	// xBusy не покрывает удерживаемый запрос и завершение Disable.
	// Занятость другого магазина/станка сама по себе не запрещает правку инвентаря.
	xTwinRobotOperation := GVL_MAGAZINE.astPartStatus[uiTwin].xBusy
		OR GVL_MAGAZINE.astPartStatus[uiTwin].xDisablePending
		OR GVL_MAGAZINE.astAutoCommand[uiTwin].xExecute
		OR GVL_MAGAZINE.astCommand[uiTwin].xExecute
		OR ((GVL_ROBOT.Status.xBusy OR xMotionBusy)
			AND (GVL_ROBOT.Status.uiMagazineContext = uiTwin))
		OR ((GVL_CELL_MANAGER.Status.uiActiveMagazine = uiTwin)
			AND ((GVL_CELL_MANAGER.Diag.eState = E_CELL_STATE.MAGAZINE)
				OR (GVL_CELL_MANAGER.Diag.eState = E_CELL_STATE.RELEASE_MAGAZINE)));
	// Для обмена важна занятость только этого магазина. Точка и состояние
	// интерфейса робота после инициализации могут быть неизвестны.
	xTwinRobotSwapWindow := NOT xTwinRobotOperation;
	xTwinOtherLoaded := FALSE;
	IF (GVL_TWO_PALLET.astStatus[uiTwin].uiRobotPallet >= UINT#1)
		AND (GVL_TWO_PALLET.astStatus[uiTwin].uiRobotPallet <= UINT#2) THEN
		uiTwinPallet := UINT#3 - GVL_TWO_PALLET.astStatus[uiTwin].uiRobotPallet;
		xTwinOtherLoaded := GVL_TWO_PALLET.astStore[uiTwin].axLoaded[uiTwinPallet];
	END_IF;
	// Finished удерживает цикл в ожидании даже до подтверждения загрузки второй палеты.
	// Подтверждение, разрешение автообмена и готовность зоны отдельно разрешают движение.
	axTwinAutoSwapPending[uiTwin] := (GVL_TWO_PALLET.uiMode = UINT#1)
		AND GVL_CELL_MANAGER.Status.xRunning
		AND NOT GVL_CELL_MANAGER.Status.xStopPending
		AND NOT GVL_CELL_CONTROL.xStop
		AND NOT GVL_CELL_CONTROL.xManual
		AND GVL_MAGAZINE.astPartStatus[uiTwin].xFinished
		AND NOT astTwinCommand[uiTwin].xDisable
		AND NOT astTwinCommand[uiTwin].xStop;
	uiTwinRobotPalletBefore := GVL_TWO_PALLET.astStatus[uiTwin].uiRobotPallet;
	TWIN[uiTwin](
		xSelected := GVL_TWO_PALLET.uiMode = 1,
		xManual := GVL_CELL_CONTROL.xManual AND NOT GVL_CELL_MANAGER.Status.xRunning,
		xSafe := CELL_SAFETY.Status.xReady AND NOT GVL_CELL_CONTROL.xGlobalError AND NOT GVL_HMI.xIoEmergencyStopActive
			AND CELL_SAFETY.astEnclosureDoorStatus[uiTwin * 2 - 1].xLocked
			AND CELL_SAFETY.astEnclosureDoorStatus[uiTwin * 2].xLocked
			AND NOT CELL_SAFETY.astEnclosureDoorStatus[uiTwin * 2 - 1].xUnlockOutput
			AND NOT CELL_SAFETY.astEnclosureDoorStatus[uiTwin * 2].xUnlockOutput,
		xRobotSwapWindow := xTwinRobotSwapWindow,
		xRobotOperation := xTwinRobotOperation,
		xPointsConfigured := axMagazinePointsReady[uiTwin],
		xRobotGeometryReady := NOT GVL_HMI.xModbusMode AND axMagazinePointsReady[uiTwin],
		xRobotMagazineReady := GVL_MAGAZINE.astPartStatus[uiTwin].xEnableCheckNoError
			AND GVL_MAGAZINE.astPartStatus[uiTwin].xEnableCheckGeometry,
		xConnection := xHmiConnectionAlive,
		xStopRequest := GVL_CELL_CONTROL.xStop OR xIoManualActive OR GVL_HMI.astMagazineCommand[uiTwin].xStop OR GVL_TWO_PALLET.xModeChanged,
		xAutoSwap := axTwinAutoSwapPending[uiTwin] AND xTwinAutoSwapEnabled AND xTwinOtherLoaded,
		xOtherLoaded := xTwinOtherLoaded,
		xActivePalletEditAllowed := NOT xTwinRobotOperation,
		xConfigurationChanged := axTwinConfigurationChanged[uiTwin],
        xIoPneumaticOverride := axIoMagazineInvalidated[uiTwin],
		xExternalCommandRejected := axTwinExternalCommandRejected[uiTwin],
		Command := astTwinCommand[uiTwin],
		Config := GVL_TWO_PALLET.astActiveConfig[uiTwin], Input := GVL_TWO_PALLET.astInput[uiTwin],
		Status => GVL_TWO_PALLET.astStatus[uiTwin],
		Diag => GVL_TWO_PALLET.astDiag[uiTwin],
		Error => GVL_TWO_PALLET.astError[uiTwin],
		Output => GVL_TWO_PALLET.astOutput[uiTwin]);
    axIoMagazineInvalidated[uiTwin] := FALSE;
	// Блокировка относится только к этому магазину и удерживается до полного
	// окончания механического обмена, включая последний скан Completed.
	axTwinMagazineExchangeInProgress[uiTwin] := GVL_TWO_PALLET.astStatus[uiTwin].xBusy
		OR GVL_TWO_PALLET.astStatus[uiTwin].xCompleted;
	GVL_TWO_PALLET.astStatus[uiTwin].xAutoSwapEnabled := xTwinAutoSwapEnabled;
	// После Stop/Disable или аварии ожидание обмена не удерживает планировщик.
	axTwinAutoSwapPending[uiTwin] := axTwinAutoSwapPending[uiTwin]
		AND NOT GVL_TWO_PALLET.astStatus[uiTwin].xError;
	axTwinConfigurationChanged[uiTwin] := FALSE;
	axTwinExternalCommandRejected[uiTwin] := FALSE;
	IF GVL_TWO_PALLET.astOutput[uiTwin].xTeachOperator THEN
		IF GVL_CELL_SETTINGS.eTestEnvironment = E_CELL_TEST_ENVIRONMENT.SIMULATION THEN
			GVL_TWO_PALLET.astSimulationConfig[uiTwin].lrExchange := GVL_TWO_PALLET.astInput[uiTwin].lrPosition;
		ELSE
			GVL_TWO_PALLET.astConfig[uiTwin].lrExchange := GVL_TWO_PALLET.astInput[uiTwin].lrPosition;
		END_IF;
		axTwinConfigurationChanged[uiTwin] := TRUE;
	END_IF;
	IF GVL_TWO_PALLET.astOutput[uiTwin].xTeachWork THEN
		IF GVL_TWO_PALLET.astStatus[uiTwin].uiSelected = UINT#1 THEN
			IF GVL_CELL_SETTINGS.eTestEnvironment = E_CELL_TEST_ENVIRONMENT.SIMULATION THEN
				GVL_TWO_PALLET.astSimulationConfig[uiTwin].lrWorkP1 := GVL_TWO_PALLET.astInput[uiTwin].lrPosition;
			ELSE
				GVL_TWO_PALLET.astConfig[uiTwin].lrWorkP1 := GVL_TWO_PALLET.astInput[uiTwin].lrPosition;
			END_IF;
		ELSIF GVL_TWO_PALLET.astStatus[uiTwin].uiSelected = UINT#2 THEN
			IF GVL_CELL_SETTINGS.eTestEnvironment = E_CELL_TEST_ENVIRONMENT.SIMULATION THEN
				GVL_TWO_PALLET.astSimulationConfig[uiTwin].lrWorkP2 := GVL_TWO_PALLET.astInput[uiTwin].lrPosition;
			ELSE
				GVL_TWO_PALLET.astConfig[uiTwin].lrWorkP2 := GVL_TWO_PALLET.astInput[uiTwin].lrPosition;
			END_IF;
		END_IF;
		axTwinConfigurationChanged[uiTwin] := TRUE;
	END_IF;
	// RunCellControl ниже должен видеть запрет уже в скане начала обмена.
	IF GVL_TWO_PALLET.uiMode = 1 THEN
		GVL_MAGAZINE.astStatus[uiTwin].xReady := GVL_MAGAZINE.astPartStatus[uiTwin].xReady
			AND GVL_TWO_PALLET.astStatus[uiTwin].xReady;
		GVL_MAGAZINE.astStatus[uiTwin].xBusy := GVL_MAGAZINE.astPartStatus[uiTwin].xBusy
			OR GVL_TWO_PALLET.astStatus[uiTwin].xBusy;
		GVL_MAGAZINE.astStatus[uiTwin].xEnabled := GVL_TWO_PALLET.astStatus[uiTwin].xEnabled;
	END_IF;
	IF GVL_TWO_PALLET.astStatus[uiTwin].xCompleted THEN
		GVL_TWO_PALLET.astStore[uiTwin].axLoaded[1] := FALSE;
		GVL_TWO_PALLET.astStore[uiTwin].axLoaded[2] := FALSE;
		axMagazineInventoryChanged[uiTwin] := TRUE;
	END_IF;
	// Ручное восстановление может сменить учётную роль без команды обмена.
	IF uiTwinRobotPalletBefore <> GVL_TWO_PALLET.astStatus[uiTwin].uiRobotPallet THEN
		GVL_TWO_PALLET.astStore[uiTwin].axLoaded[1] := FALSE;
		GVL_TWO_PALLET.astStore[uiTwin].axLoaded[2] := FALSE;
		axMagazineInventoryChanged[uiTwin] := TRUE;
	END_IF;
	// Ручная смена расходует прежнее подтверждение уже при принятии команды.
	IF astTwinCommand[uiTwin].xSwap AND GVL_TWO_PALLET.astStatus[uiTwin].xCommandAccepted THEN
		GVL_TWO_PALLET.astStore[uiTwin].axLoaded[1] := FALSE;
		GVL_TWO_PALLET.astStore[uiTwin].axLoaded[2] := FALSE;
	END_IF;
	IF (uiTwinRequestResult = 2) AND (stTwinRequest.uiMagazine = uiTwin)
		AND (((stTwinRequest.uiCommand >= 1) AND (stTwinRequest.uiCommand <= 19))
			OR ((stTwinRequest.uiCommand >= 25) AND (stTwinRequest.uiCommand <= 32)))
		AND GVL_TWO_PALLET.astStatus[uiTwin].xCommandAccepted THEN uiTwinRequestResult := 1; END_IF;
END_FOR;

IF xTwinInventoryCommand THEN
	uiTwin := stTwinRequest.uiMagazine;
	uiTwinPallet := stTwinRequest.uiValue;
	IF stTwinRequest.uiCommand = UINT#24 THEN
		IF GVL_TWO_PALLET.astStatus[uiTwin].xConfigAllowed
			AND stTwinRequest.Config.xSignalPatternsConfigured
			AND TWIN[uiTwin].IsSignalConfigurationValid(
				uiP1Signals := stTwinRequest.Config.uiP1Signals,
				uiP2Signals := stTwinRequest.Config.uiP2Signals) THEN
			IF GVL_CELL_SETTINGS.eTestEnvironment = E_CELL_TEST_ENVIRONMENT.SIMULATION THEN
				GVL_TWO_PALLET.astSimulationConfig[uiTwin] := stTwinRequest.Config;
			ELSE
				GVL_TWO_PALLET.astConfig[uiTwin] := stTwinRequest.Config;
			END_IF;
			axTwinConfigurationChanged[uiTwin] := TRUE;
			uiTwinRequestResult := UINT#1;
		END_IF;
	ELSIF ((uiTwinPallet = 1) AND GVL_TWO_PALLET.astStatus[uiTwin].xEdit1Allowed)
		OR ((uiTwinPallet = 2) AND GVL_TWO_PALLET.astStatus[uiTwin].xEdit2Allowed) THEN
		CASE stTwinRequest.uiCommand OF
			20:
				IF GVL_TWO_PALLET.astStatus[uiTwin].xLoadAllowed
					AND (uiTwinPallet <> GVL_TWO_PALLET.astStatus[uiTwin].uiRobotPallet) THEN
					GVL_TWO_PALLET.astStore[uiTwin].axLoaded[uiTwinPallet] := TRUE;
					uiTwinRequestResult := 1;
				END_IF;
			21, 22:
				FOR uiTwinSlot := 1 TO 96 DO
					GVL_TWO_PALLET.astStore[uiTwin].astPallet[uiTwinPallet].aSlots[uiTwinSlot].xInPosition := stTwinRequest.uiCommand = 22;
					GVL_TWO_PALLET.astStore[uiTwin].astPallet[uiTwinPallet].aSlots[uiTwinSlot].eDetailType := E_DETAIL_TYPE.NONE;
					GVL_TWO_PALLET.astStore[uiTwin].astPallet[uiTwinPallet].aSlots[uiTwinSlot].uiProductType := 0;
					IF stTwinRequest.uiCommand = 22 THEN
						GVL_TWO_PALLET.astStore[uiTwin].astPallet[uiTwinPallet].aSlots[uiTwinSlot].eDetailType := E_DETAIL_TYPE.BLANK;
						GVL_TWO_PALLET.astStore[uiTwin].astPallet[uiTwinPallet].aSlots[uiTwinSlot].uiProductType := GVL_MULTI_TYPE.Config.auiSlotType[uiTwinSlot];
					END_IF;
				END_FOR;
				GVL_TWO_PALLET.astStore[uiTwin].axLoaded[uiTwinPallet] := FALSE; uiTwinRequestResult := 1;
			23:
				IF (stTwinRequest.uiSlot >= 1) AND (stTwinRequest.uiSlot <= 96) AND (stTwinRequest.uiContent <= 2)
					AND ((stTwinRequest.uiContent = 0) OR ((stTwinRequest.uiProductType >= 1) AND (stTwinRequest.uiProductType <= GVL_MULTI_TYPE.Config.uiTypeCount))) THEN
					uiTwinSlot := stTwinRequest.uiSlot;
					GVL_TWO_PALLET.astStore[uiTwin].astPallet[uiTwinPallet].aSlots[uiTwinSlot].xInPosition := stTwinRequest.uiContent <> 0;
					CASE stTwinRequest.uiContent OF
						0: GVL_TWO_PALLET.astStore[uiTwin].astPallet[uiTwinPallet].aSlots[uiTwinSlot].eDetailType := E_DETAIL_TYPE.NONE;
						1: GVL_TWO_PALLET.astStore[uiTwin].astPallet[uiTwinPallet].aSlots[uiTwinSlot].eDetailType := E_DETAIL_TYPE.BLANK;
						2: GVL_TWO_PALLET.astStore[uiTwin].astPallet[uiTwinPallet].aSlots[uiTwinSlot].eDetailType := E_DETAIL_TYPE.DETAIL;
					END_CASE;
					GVL_TWO_PALLET.astStore[uiTwin].astPallet[uiTwinPallet].aSlots[uiTwinSlot].uiProductType := stTwinRequest.uiProductType;
					GVL_TWO_PALLET.astStore[uiTwin].axLoaded[uiTwinPallet] := FALSE; uiTwinRequestResult := 1;
				END_IF;
		END_CASE;
		// Загрузка/редактирование палеты у оператора не отменяет завершение рабочей.
		IF (uiTwinRequestResult = UINT#1)
			AND (stTwinRequest.uiCommand >= UINT#21)
			AND (stTwinRequest.uiCommand <= UINT#23)
			AND (uiTwinPallet = GVL_TWO_PALLET.astStatus[uiTwin].uiRobotPallet) THEN
			axMagazineInventoryChanged[uiTwin] := TRUE;
		END_IF;
	END_IF;
END_IF;
IF uiTwinRequestResult <> 0 THEN
	GVL_HMI.uiTwinResult := uiTwinRequestResult;
	GVL_HMI.udiTwinAckSeq := udiTwinSnapshot;
	IF uiTwinRequestResult <> 1 THEN
		uiTwin := LIMIT(UINT#1, stTwinRequest.uiMagazine, UINT#2);
		// Команды механизма 1..19 и 25..28 уже формируют предупреждение внутри FB в этом же скане.
		IF GVL_TWO_PALLET.auiCommand[uiTwin] <> stTwinRequest.uiCommand THEN
			axTwinExternalCommandRejected[uiTwin] := TRUE;
		END_IF;
	END_IF;
END_IF;

GVL_CELL_SETTINGS.MagazineRows := 12;
GVL_CELL_SETTINGS.MagazineColumns := 10;
IF GVL_TWO_PALLET.uiMode = 1 THEN GVL_CELL_SETTINGS.MagazineRows := 12; GVL_CELL_SETTINGS.MagazineColumns := 8; END_IF;
GVL_HMI.MagazineRows := GVL_CELL_SETTINGS.MagazineRows;
GVL_HMI.MagazineColumns := GVL_CELL_SETTINGS.MagazineColumns;
FOR uiTwin := 1 TO 2 DO
	IF GVL_TWO_PALLET.uiMode = 1 THEN
		uiTwinPallet := GVL_TWO_PALLET.astStatus[uiTwin].uiRobotPallet;
		IF (uiTwinPallet < UINT#1) OR (uiTwinPallet > UINT#2) THEN
			uiTwinPallet := UINT#1;
		END_IF;
		GVL_DETAIL.astMagazine[uiTwin] := GVL_TWO_PALLET.astStore[uiTwin].astPallet[uiTwinPallet];
	END_IF;
END_FOR;
END_METHOD

METHOD PRIVATE RunCellControl
// Выключенные станки, магазины и ГК не требуют настройки своих точек.
// Общая безопасная точка обязательна при любом составе автоцикла.
xCellPointsReady := GVL_POINT.Points[E_POINT_NAME.HOME_SAFETY].xConfigured;
FOR uiMachine := UINT#1 TO UINT#3 DO
	IF GVL_MACHINE.Status[uiMachine].xEnabled THEN
		xCellPointsReady := xCellPointsReady AND axMachinePointsReady[uiMachine];
	END_IF;
END_FOR;
FOR uiMagazine := UINT#1 TO UINT#2 DO
	IF GVL_MAGAZINE.astStatus[uiMagazine].xEnabled THEN
		xCellPointsReady := xCellPointsReady AND axMagazinePointsReady[uiMagazine];
	END_IF;
	IF GVL_GEOMETRY_CONTROL.astStatus[uiMagazine].xEnabled THEN
		xCellPointsReady := xCellPointsReady
			AND GVL_GEOMETRY_CONTROL.astStatus[uiMagazine].xConfigured;
	END_IF;
END_FOR;

uiMagazine := GVL_CELL_MANAGER.Status.uiActiveMagazine;
IF (uiMagazine < UINT#1) OR (uiMagazine > UINT#2) THEN
	uiMagazine := UINT#1;
END_IF;

TYPE_CONFIG(
	xTestInitialize := xTestInitializePulse,
	stTestScenario := GVL_HMI.stTestScenario,
	Command := GVL_HMI.stMultiType.Command,
	xCellRunning := GVL_CELL_MANAGER.Status.xRunning,
	xMotionBusy := xMotionBusy,
	stRobotStatus := GVL_ROBOT.Status,
	astMagazineStatus := GVL_MAGAZINE.astStatus,
	astMachineStatus := GVL_MACHINE.Status,
	uiRows := GVL_CELL_SETTINGS.MagazineRows,
	uiColumns := GVL_CELL_SETTINGS.MagazineColumns,
	Config => GVL_MULTI_TYPE.Config,
	Status => GVL_MULTI_TYPE.ConfigStatus
);

CELL_MANAGER(
	axMagazineAutoSwapPending := axTwinAutoSwapPending,
	axMagazineExchangeInProgress := axTwinMagazineExchangeInProgress,
	xMagazineExchangeActive := (GVL_TWO_PALLET.uiMode = 1) AND (
		GVL_TWO_PALLET.astStatus[1].xBusy OR GVL_TWO_PALLET.astStatus[2].xBusy
		OR GVL_TWO_PALLET.astStatus[1].xCompleted OR GVL_TWO_PALLET.astStatus[2].xCompleted),
	xStart := GVL_CELL_CONTROL.xStart,
	xStop := GVL_CELL_CONTROL.xStop,
	xTestAbort := xTestAbortActive,
	xResetRequest := GVL_HMI.xCellReset,
	xReset := GVL_CELL_CONTROL.xReset,
	xOperatorChoice := GVL_HMI.xCellOperatorChoice,
	xOperatorCancel := GVL_HMI.xCellOperatorCancel,
	uiOperatorChoice := GVL_HMI.uiCellOperatorChoice,
	xManual := GVL_CELL_CONTROL.xManual,
	xIoManual := xIoManualActive,
	uiModeRejectReason := uiCellModeRejectReason,
	xSettingsRejected := xCellSettingRejected,
	xIoOverrideRejected := xIoOverrideRejected,
    xIoDoRejected := xIoDoRejected,
    xIoEmergencyResetRejected := xIoEmergencyResetRejected,
    xIoEmergencyStopActive := GVL_HMI.xIoEmergencyStopActive,
	xGlobalError := GVL_CELL_CONTROL.xGlobalError,
	xSafetyReady := CELL_SAFETY.Status.xReady,
	xDrivesReady := xDrivesReady,
	xMotionBusy := xMotionBusy,
	xRobotInterfaceReady := xRobotInterfaceReady,
	lrRobotActualX := lrRobotActualX,
	lrRobotActualY := lrRobotActualY,
	lrRobotActualZ := lrRobotActualZ,
	stSafetyHomePoint := GVL_POINT.Points[E_POINT_NAME.HOME_SAFETY],
	lrSafetyHomeToleranceX := GVL_CELL_SETTINGS.lrSafetyHomeToleranceX,
	lrSafetyHomeToleranceY := GVL_CELL_SETTINGS.lrSafetyHomeToleranceY,
	lrSafetyHomeToleranceZ := GVL_CELL_SETTINGS.lrSafetyHomeToleranceZ,
	lrStoppedPoseTolerance := GVL_CELL_SETTINGS.lrStoppedPoseTolerance,
	Config := GVL_MULTI_TYPE.Config,
	xConfigurationValid := GVL_MULTI_TYPE.ConfigStatus.xConfigurationValid,
	xPointsConfigured := xCellPointsReady,
	stRobotStatus := GVL_ROBOT.Status,
	astMagazineStatus := GVL_MAGAZINE.astStatus,
	astMachineStatus := GVL_MACHINE.Status,
	astMachineDiag := GVL_MACHINE.Diag,
	FaultRequest := stCellFaultRequest,
	Command => GVL_CELL_MANAGER.Command,
	Status => GVL_CELL_MANAGER.Status,
	Diag => GVL_CELL_MANAGER.Diag,
	Error => GVL_CELL_MANAGER.Error,
	CycleStatus => GVL_MULTI_TYPE.CycleStatus
);

// Сначала снимаем команды обоих владельцев, затем маршрутизируем единственную
// команду менеджера выбранному магазину.
// Общий Disable ячейки не отключает независимо включённые магазины.
FOR uiMagazine := UINT#1 TO UINT#2 DO
	GVL_MAGAZINE.astAutoCommand[uiMagazine].xEnable := FALSE;
	GVL_MAGAZINE.astAutoCommand[uiMagazine].xDisable := FALSE;
	GVL_MAGAZINE.astAutoCommand[uiMagazine].xExecute := FALSE;
	GVL_MAGAZINE.astAutoCommand[uiMagazine].xStop := FALSE;
	GVL_MAGAZINE.astAutoCommand[uiMagazine].eOperation := E_MAGAZINE_OPERATION.NONE;
	GVL_MAGAZINE.astAutoCommand[uiMagazine].iTakeSlot := SINT#0;
	GVL_MAGAZINE.astAutoCommand[uiMagazine].iPutSlot := SINT#0;
END_FOR;
IF (GVL_CELL_MANAGER.Status.uiActiveMagazine >= UINT#1)
AND (GVL_CELL_MANAGER.Status.uiActiveMagazine <= UINT#2) THEN
	GVL_MAGAZINE.astAutoCommand[GVL_CELL_MANAGER.Status.uiActiveMagazine] :=
		GVL_CELL_MANAGER.Command.stMagazine;
	GVL_MAGAZINE.astAutoCommand[GVL_CELL_MANAGER.Status.uiActiveMagazine].xEnable := FALSE;
END_IF;
END_METHOD

METHOD PRIVATE RunTestControl
// Test environment is independent from the robot control interface.
rtTestEnvironmentApply(CLK := GVL_HMI.xTestEnvironmentApply);
rtTestSpeedProfileApply(CLK := GVL_HMI.xTestSpeedProfileApply);
rtTestScenarioApply(CLK := GVL_HMI.xTestScenarioApply);
xTestInitializePulse := FALSE;
xTestAbortActive := GVL_HMI.xTestAbort
	AND GVL_HMI.xTestSessionActive
	AND (GVL_CELL_SETTINGS.eTestEnvironment = E_CELL_TEST_ENVIRONMENT.SIMULATION);

xTestStable := NOT GVL_CELL_MANAGER.Status.xRunning
	AND NOT GVL_ROBOT.Status.xBusy
	AND NOT GVL_MAGAZINE.astStatus[1].xBusy
	AND NOT GVL_MAGAZINE.astStatus[2].xBusy
	AND NOT GVL_TWO_PALLET.astInput[1].xPowered
	AND NOT GVL_TWO_PALLET.astInput[2].xPowered
	AND NOT xMotionBusy
	AND NOT SIMULATION_DYNAMICS.xBusy;
FOR uiTestIndex := UINT#1 TO UINT#3 DO
	xTestStable := xTestStable
		AND NOT GVL_MACHINE.Status[uiTestIndex].xBusy
		AND NOT GVL_MACHINE.Status[uiTestIndex].xProcessing;
END_FOR;

GVL_HMI.xTestEnvironmentChangeAllowed := xTestStable;
GVL_HMI.xTestScenarioApplyAllowed := xTestStable
	AND (GVL_TWO_PALLET.uiMode = 0) // Existing scenarios describe static 120-slot magazines
	AND GVL_HMI.xTestSessionActive
	AND (GVL_CELL_SETTINGS.eTestEnvironment <> E_CELL_TEST_ENVIRONMENT.NORMAL)
	AND ((GVL_CELL_SETTINGS.eTestEnvironment <> E_CELL_TEST_ENVIRONMENT.SIMULATION)
		OR NOT GVL_ROBOT_MODBUS.xModeActive
		OR GVL_ROBOT_MODBUS.Status.xSimulatorActive);
// Старые OPC UA поля сохранены для совместимости; физический ключ исключён.
GVL_HMI.xSc500BenchKeyActive := FALSE;

IF rtTestEnvironmentApply.Q THEN
	GVL_HMI.uiTestRejectReason := UINT#0;
	IF NOT GVL_HMI.xTestEnvironmentChangeAllowed THEN
		GVL_HMI.uiTestRejectReason := UINT#1; // equipment is not idle
	ELSIF GVL_HMI.uiTestEnvironmentRequest > UINT#2 THEN
		GVL_HMI.uiTestRejectReason := UINT#2; // invalid environment
	ELSIF (GVL_HMI.uiTestEnvironmentRequest = UINT#2)
	AND NOT GVL_ROBOT_MODBUS.xModeActive THEN
		GVL_HMI.uiTestRejectReason := UINT#3; // bench requires Modbus
	ELSIF (GVL_HMI.uiTestEnvironmentRequest = UINT#1)
	AND GVL_ROBOT_MODBUS.xModeActive
	AND NOT GVL_ROBOT_MODBUS.Status.xSimulatorActive THEN
		GVL_HMI.uiTestRejectReason := UINT#4; // Python simulator marker missing
	ELSE
		CASE GVL_HMI.uiTestEnvironmentRequest OF
			UINT#0: GVL_CELL_SETTINGS.eTestEnvironment := E_CELL_TEST_ENVIRONMENT.NORMAL;
			UINT#1: GVL_CELL_SETTINGS.eTestEnvironment := E_CELL_TEST_ENVIRONMENT.SIMULATION;
			UINT#2: GVL_CELL_SETTINGS.eTestEnvironment := E_CELL_TEST_ENVIRONMENT.SC500_BENCH;
		END_CASE;
		IF GVL_CELL_SETTINGS.eTestEnvironment = E_CELL_TEST_ENVIRONMENT.NORMAL THEN
			GVL_CELL_SETTINGS.xErrorSimulationEnabled := FALSE;
		END_IF;
		GVL_CELL_SETTINGS.eTestSpeedProfile := E_TEST_SPEED_PROFILE.REALTIME;
	END_IF;
END_IF;

IF rtTestSpeedProfileApply.Q THEN
	GVL_HMI.uiTestRejectReason := UINT#0;
	IF (GVL_HMI.uiTestSpeedProfileRequest <= UINT#1)
	AND (GVL_CELL_SETTINGS.eTestEnvironment = E_CELL_TEST_ENVIRONMENT.SIMULATION) THEN
		IF GVL_HMI.uiTestSpeedProfileRequest = UINT#1 THEN
			GVL_CELL_SETTINGS.eTestSpeedProfile := E_TEST_SPEED_PROFILE.FAST;
			// В Modbus профиль по-прежнему владеет коэффициентом внешней модели.
			// В SoftMotion коэффициент задаёт ползунок, а применение выполняется
			// отдельной транзакцией только на границе следующего теста.
			IF GVL_ROBOT_MODBUS.xModeActive THEN
				GVL_CELL_SETTINGS.uiSimulationTimeFactor := UINT#250;
			END_IF;
		ELSE
			GVL_CELL_SETTINGS.eTestSpeedProfile := E_TEST_SPEED_PROFILE.REALTIME;
			IF GVL_ROBOT_MODBUS.xModeActive THEN
				GVL_CELL_SETTINGS.uiSimulationTimeFactor := UINT#1;
			END_IF;
		END_IF;
		GVL_HMI.uiSimulationTimeFactor := GVL_CELL_SETTINGS.uiSimulationTimeFactor;
	ELSE
		GVL_HMI.uiTestRejectReason := UINT#5; // speed profile is simulation-only
	END_IF;
END_IF;

IF rtTestScenarioApply.Q THEN
	GVL_HMI.uiTestScenarioResult := UINT#0;
	xTestScenarioValid := GVL_HMI.stTestScenario.udiLoadSeq <> UDINT#0
		AND (GVL_HMI.stTestScenario.uiTypeCount >= UINT#1)
		AND (GVL_HMI.stTestScenario.uiTypeCount <= UINT#3);
	FOR uiTestIndex := UINT#1 TO UINT#3 DO
		xTestScenarioValid := xTestScenarioValid
			AND (GVL_HMI.stTestScenario.auiMachineState[uiTestIndex] <= UINT#3)
			AND (GVL_HMI.stTestScenario.auiMachineType[uiTestIndex] >= UINT#1)
			AND (GVL_HMI.stTestScenario.auiMachineType[uiTestIndex]
				<= GVL_HMI.stTestScenario.uiTypeCount);
	END_FOR;
	FOR uiTestIndex := UINT#1 TO UINT#120 DO
		xTestScenarioValid := xTestScenarioValid
			AND (GVL_HMI.stTestScenario.auiSlotType[uiTestIndex] >= UINT#1)
			AND (GVL_HMI.stTestScenario.auiSlotType[uiTestIndex]
				<= GVL_HMI.stTestScenario.uiTypeCount);
		FOR uiTestMagazine := UINT#1 TO UINT#2 DO
			xTestScenarioValid := xTestScenarioValid
				AND (GVL_HMI.stTestScenario.aauiSlotContent[uiTestMagazine, uiTestIndex] <= UINT#2);
		END_FOR;
	END_FOR;
	uiTestFaultOwnerCount := UINT#0;
	IF GVL_HMI.stTestScenario.dwCellFaultMask <> DWORD#0 THEN
		uiTestFaultOwnerCount := uiTestFaultOwnerCount + UINT#1;
	END_IF;
	IF GVL_HMI.stTestScenario.dwRobotFaultMask <> DWORD#0 THEN
		uiTestFaultOwnerCount := uiTestFaultOwnerCount + UINT#1;
	END_IF;
	FOR uiTestMagazine := UINT#1 TO UINT#2 DO
		IF GVL_HMI.stTestScenario.adwMagazineFaultMask[uiTestMagazine] <> DWORD#0 THEN
			uiTestFaultOwnerCount := uiTestFaultOwnerCount + UINT#1;
		END_IF;
		xTestScenarioValid := xTestScenarioValid
			AND (GVL_HMI.stTestScenario.adwMagazineFaultMask[uiTestMagazine] <= DWORD#16#0000_003F);
	END_FOR;
	FOR uiTestIndex := UINT#1 TO UINT#3 DO
		IF GVL_HMI.stTestScenario.adwMachineFaultMask[uiTestIndex] <> DWORD#0 THEN
			uiTestFaultOwnerCount := uiTestFaultOwnerCount + UINT#1;
		END_IF;
		xTestScenarioValid := xTestScenarioValid
			AND (GVL_HMI.stTestScenario.adwMachineFaultMask[uiTestIndex] <= DWORD#16#0000_07FF);
	END_FOR;
	xTestScenarioValid := xTestScenarioValid
		AND (uiTestFaultOwnerCount <= UINT#1)
		AND (GVL_HMI.stTestScenario.dwCellFaultMask <= DWORD#16#0000_0001)
		AND (GVL_HMI.stTestScenario.dwRobotFaultMask <= DWORD#16#0000_01FF)
		AND (GVL_HMI.stTestScenario.auiGripperContent[1] <= UINT#1)
		AND ((GVL_HMI.stTestScenario.auiGripperContent[1] = UINT#0)
			= (GVL_HMI.stTestScenario.auiGripperType[1] = UINT#0))
		AND (GVL_HMI.stTestScenario.auiGripperType[1]
			<= GVL_HMI.stTestScenario.uiTypeCount)
		AND ((GVL_HMI.stTestScenario.auiGripperContent[2] = UINT#0)
			OR (GVL_HMI.stTestScenario.auiGripperContent[2] = UINT#2))
		AND ((GVL_HMI.stTestScenario.auiGripperContent[2] = UINT#0)
			= (GVL_HMI.stTestScenario.auiGripperType[2] = UINT#0))
		AND (GVL_HMI.stTestScenario.auiGripperType[2]
			<= GVL_HMI.stTestScenario.uiTypeCount);

	IF NOT GVL_HMI.xTestScenarioApplyAllowed THEN
		GVL_HMI.uiTestScenarioResult := UINT#1;
	ELSIF NOT xTestScenarioValid OR (GVL_HMI.stTestScenario.uiOrientation > UINT#1) THEN
		GVL_HMI.uiTestScenarioResult := UINT#2;
	ELSE
		FOR uiTestMagazine := UINT#1 TO UINT#2 DO
			FOR uiTestIndex := UINT#1 TO UINT#120 DO
				GVL_DETAIL.astMagazine[uiTestMagazine].aSlots[uiTestIndex].xInPosition :=
					GVL_HMI.stTestScenario.aauiSlotContent[uiTestMagazine, uiTestIndex] <> UINT#0;
				CASE GVL_HMI.stTestScenario.aauiSlotContent[uiTestMagazine, uiTestIndex] OF
					UINT#1: GVL_DETAIL.astMagazine[uiTestMagazine].aSlots[uiTestIndex].eDetailType := E_DETAIL_TYPE.BLANK;
					UINT#2: GVL_DETAIL.astMagazine[uiTestMagazine].aSlots[uiTestIndex].eDetailType := E_DETAIL_TYPE.DETAIL;
				ELSE
					GVL_DETAIL.astMagazine[uiTestMagazine].aSlots[uiTestIndex].eDetailType := E_DETAIL_TYPE.NONE;
				END_CASE;
				IF GVL_HMI.stTestScenario.aauiSlotContent[uiTestMagazine, uiTestIndex] = UINT#0 THEN
					GVL_DETAIL.astMagazine[uiTestMagazine].aSlots[uiTestIndex].uiProductType := UINT#0;
				ELSE
					GVL_DETAIL.astMagazine[uiTestMagazine].aSlots[uiTestIndex].uiProductType :=
						GVL_HMI.stTestScenario.auiSlotType[uiTestIndex];
				END_IF;
			END_FOR;
			adwTestMagazineFaultMask[uiTestMagazine] :=
				GVL_HMI.stTestScenario.adwMagazineFaultMask[uiTestMagazine];
		END_FOR;
		// Начальные инъекции: маски переводятся в существующий диагностический
		// контракт, а не обходят владельцев ошибок.
		axHmiInternalPulse[13] :=
			(GVL_HMI.stTestScenario.dwCellFaultMask AND DWORD#16#0000_0001) <> DWORD#0;
		axHmiInternalPulse[12] :=
			(GVL_HMI.stTestScenario.dwRobotFaultMask AND DWORD#16#0000_0001) <> DWORD#0;
		GVL_HMI.xSimGripper1Fault :=
			(GVL_HMI.stTestScenario.dwRobotFaultMask AND DWORD#16#0000_0002) <> DWORD#0;
		GVL_HMI.xSimGripper2Fault :=
			(GVL_HMI.stTestScenario.dwRobotFaultMask AND DWORD#16#0000_0004) <> DWORD#0;
		GVL_HMI.xSimGripperRotationFault :=
			(GVL_HMI.stTestScenario.dwRobotFaultMask AND DWORD#16#0000_0008) <> DWORD#0;
		GVL_HMI.xSimGripperGlobalFault :=
			(GVL_HMI.stTestScenario.dwRobotFaultMask AND DWORD#16#0000_0010) <> DWORD#0;
		axHmiInternalPulse[14] :=
			(GVL_HMI.stTestScenario.dwRobotFaultMask AND DWORD#16#0000_0020) <> DWORD#0;
		axHmiInternalPulse[15] :=
			(GVL_HMI.stTestScenario.dwRobotFaultMask AND DWORD#16#0000_0040) <> DWORD#0;
		axHmiInternalPulse[16] :=
			(GVL_HMI.stTestScenario.dwRobotFaultMask AND DWORD#16#0000_0080) <> DWORD#0;
		axHmiInternalPulse[17] :=
			(GVL_HMI.stTestScenario.dwRobotFaultMask AND DWORD#16#0000_0100) <> DWORD#0;
		axHmiInternalPulse[18] :=
			(GVL_HMI.stTestScenario.adwMagazineFaultMask[1] AND DWORD#16#0000_0001) <> DWORD#0;
		axHmiInternalPulse[19] :=
			(GVL_HMI.stTestScenario.adwMagazineFaultMask[1] AND DWORD#16#0000_0002) <> DWORD#0;
		axHmiInternalPulse[20] :=
			(GVL_HMI.stTestScenario.adwMagazineFaultMask[1] AND DWORD#16#0000_0004) <> DWORD#0;
		axHmiInternalPulse[21] :=
			(GVL_HMI.stTestScenario.adwMagazineFaultMask[1] AND DWORD#16#0000_0008) <> DWORD#0;
		axHmiInternalPulse[22] :=
			(GVL_HMI.stTestScenario.adwMagazineFaultMask[1] AND DWORD#16#0000_0010) <> DWORD#0;
		axHmiInternalPulse[23] :=
			(GVL_HMI.stTestScenario.adwMagazineFaultMask[1] AND DWORD#16#0000_0020) <> DWORD#0;
		FOR uiTestIndex := UINT#1 TO UINT#3 DO
			GVL_HMI.axMachineSimAlarm[uiTestIndex] :=
				(GVL_HMI.stTestScenario.adwMachineFaultMask[uiTestIndex] AND DWORD#16#0000_0001) <> DWORD#0;
			GVL_HMI.axMachineSimDoorFault[uiTestIndex] :=
				(GVL_HMI.stTestScenario.adwMachineFaultMask[uiTestIndex] AND DWORD#16#0000_0002) <> DWORD#0;
			GVL_HMI.axMachineSimChuckFault[uiTestIndex] :=
				(GVL_HMI.stTestScenario.adwMachineFaultMask[uiTestIndex] AND DWORD#16#0000_0004) <> DWORD#0;
			GVL_HMI.axMachineTimeoutRobotMove[uiTestIndex] :=
				(GVL_HMI.stTestScenario.adwMachineFaultMask[uiTestIndex] AND DWORD#16#0000_0008) <> DWORD#0;
			GVL_HMI.axMachineTimeoutRobotAction[uiTestIndex] :=
				(GVL_HMI.stTestScenario.adwMachineFaultMask[uiTestIndex] AND DWORD#16#0000_0010) <> DWORD#0;
			GVL_HMI.axMachineTimeoutRobotRelease[uiTestIndex] :=
				(GVL_HMI.stTestScenario.adwMachineFaultMask[uiTestIndex] AND DWORD#16#0000_0020) <> DWORD#0;
			GVL_HMI.axMachineTimeoutDoorOpen[uiTestIndex] :=
				(GVL_HMI.stTestScenario.adwMachineFaultMask[uiTestIndex] AND DWORD#16#0000_0040) <> DWORD#0;
			GVL_HMI.axMachineTimeoutDoorClose[uiTestIndex] :=
				(GVL_HMI.stTestScenario.adwMachineFaultMask[uiTestIndex] AND DWORD#16#0000_0080) <> DWORD#0;
			GVL_HMI.axMachineTimeoutChuckOpen[uiTestIndex] :=
				(GVL_HMI.stTestScenario.adwMachineFaultMask[uiTestIndex] AND DWORD#16#0000_0100) <> DWORD#0;
			GVL_HMI.axMachineTimeoutChuckClose[uiTestIndex] :=
				(GVL_HMI.stTestScenario.adwMachineFaultMask[uiTestIndex] AND DWORD#16#0000_0200) <> DWORD#0;
			GVL_HMI.axMachineTimeoutCycleStart[uiTestIndex] :=
				(GVL_HMI.stTestScenario.adwMachineFaultMask[uiTestIndex] AND DWORD#16#0000_0400) <> DWORD#0;
		END_FOR;
		GVL_HMI.xErrorSimulationEnable :=
			(GVL_HMI.stTestScenario.dwCellFaultMask <> DWORD#0)
			OR (GVL_HMI.stTestScenario.dwRobotFaultMask <> DWORD#0)
			OR (GVL_HMI.stTestScenario.adwMagazineFaultMask[1] <> DWORD#0)
			OR (GVL_HMI.stTestScenario.adwMagazineFaultMask[2] <> DWORD#0)
			OR (GVL_HMI.stTestScenario.adwMachineFaultMask[1] <> DWORD#0)
			OR (GVL_HMI.stTestScenario.adwMachineFaultMask[2] <> DWORD#0)
			OR (GVL_HMI.stTestScenario.adwMachineFaultMask[3] <> DWORD#0);
		xTestInitializePulse := TRUE;
	END_IF;
	// Ack подтверждает обработку конкретного LoadSeq даже при отклонении.
	GVL_HMI.udiTestScenarioAckSeq := GVL_HMI.stTestScenario.udiLoadSeq;
END_IF;

GVL_HMI.uiTestEnvironmentApplied := TO_UINT(GVL_CELL_SETTINGS.eTestEnvironment);
GVL_HMI.uiTestSpeedProfileApplied := TO_UINT(GVL_CELL_SETTINGS.eTestSpeedProfile);
GVL_HMI.xSc500BenchKeyLost := FALSE;
IF GVL_CELL_SETTINGS.eTestEnvironment = E_CELL_TEST_ENVIRONMENT.SIMULATION THEN
	IF GVL_HMI.xTestSessionActive THEN
		GVL_CELL_SETTINGS.xSimulationAccelerationEnable :=
			GVL_CELL_SETTINGS.eTestSpeedProfile = E_TEST_SPEED_PROFILE.FAST;
		// Профиль владеет включением ускоренных таймеров, а сам коэффициент
		// разрешено менять с HMI прямо во время тестового движения.
		GVL_HMI.xSimulationAccelerationEnable := GVL_CELL_SETTINGS.xSimulationAccelerationEnable;
	END_IF;
ELSE
	GVL_CELL_SETTINGS.xSimulationAccelerationEnable := FALSE;
	GVL_HMI.xSimulationAccelerationEnable := FALSE;
END_IF;
END_METHOD

METHOD PRIVATE RunSignalTower
VAR
	xBlink : BOOL;
END_VAR
fbAlarmHorn(astSource := astAlarmSource, tDuration := GVL_CELL_SETTINGS.tAlarmHornDuration);
GVL_CELL_SAFETY_IO.xAlarmHornOutput := fbAlarmHorn.xSound;

// Приоритет: авария > предупреждение > работа > готовность > остановлена/не готова.
// Вызывать после RunAlarms: используются актуальные сводные состояния этого скана.
IF GVL_ALARM.Status.xAlarmActive THEN
	usiSignalTowerMode := USINT#4;
ELSIF GVL_ALARM.Status.xWarningActive THEN
	usiSignalTowerMode := USINT#3;
ELSIF GVL_CELL_MANAGER.Status.xRunning THEN
	usiSignalTowerMode := USINT#1;
ELSIF GVL_CELL_MANAGER.Status.xReadyToStart THEN
	usiSignalTowerMode := USINT#2;
ELSE
	usiSignalTowerMode := USINT#5;
END_IF;

xBlink := (usiSignalTowerMode = USINT#2) OR (usiSignalTowerMode = USINT#4);
tonSignalTowerBlink(
	IN := xBlink AND (usiSignalTowerMode = usiSignalTowerPreviousMode) AND NOT tonSignalTowerBlink.Q,
	PT := T#500MS
);
// Каждый новый режим начинается со включённой секции, без ожидания таймера.
IF (usiSignalTowerMode <> usiSignalTowerPreviousMode) OR NOT xBlink THEN
	xSignalTowerBlinkOn := TRUE;
ELSIF tonSignalTowerBlink.Q THEN
	xSignalTowerBlinkOn := NOT xSignalTowerBlinkOn;
END_IF;
usiSignalTowerPreviousMode := usiSignalTowerMode;

GVL_CELL_SAFETY_IO.xSignalTowerRedOutput := (usiSignalTowerMode = USINT#5)
	OR ((usiSignalTowerMode = USINT#4) AND xSignalTowerBlinkOn);
GVL_CELL_SAFETY_IO.xSignalTowerAmberOutput := usiSignalTowerMode = USINT#3;
GVL_CELL_SAFETY_IO.xSignalTowerGreenOutput := (usiSignalTowerMode = USINT#1)
	OR ((usiSignalTowerMode = USINT#2) AND xSignalTowerBlinkOn);
END_METHOD

METHOD PRIVATE AppendIoEvent
VAR_INPUT
    usiDirection : USINT;
    uiIndex : UINT;
    usiKind : USINT;
    xOld : BOOL;
    xNew : BOOL;
END_VAR
VAR
    uiSlot : UINT;
    sEvent : STRING(96);
END_VAR
IF NOT xIoSnapshotPublishing THEN
    GVL_HMI.udiIoJournalRevision := GVL_HMI.udiIoJournalRevision + UDINT#1;
END_IF;
// Переполнение Seq открывает новый FIFO; идентификаторы не повторяются внутри эпохи.
IF GVL_HMI.udiIoJournalSequence = UDINT#4294967295 THEN
    GVL_HMI.udiIoBootCounter := GVL_HMI.udiIoBootCounter + UDINT#1;
    IF GVL_HMI.udiIoBootCounter = UDINT#0 THEN GVL_HMI.udiIoBootCounter := UDINT#1; END_IF;
    GVL_HMI.udiIoJournalSequence := UDINT#0;
    GVL_HMI.uiIoJournalHead := UINT#0;
    GVL_HMI.uiIoJournalCount := UINT#0;
END_IF;
uiSlot := (GVL_HMI.uiIoJournalHead MOD UINT#100) + UINT#1;
GVL_HMI.udiIoJournalSequence := GVL_HMI.udiIoJournalSequence + UDINT#1;
astIoEvent[uiSlot].udiSequence := GVL_HMI.udiIoJournalSequence;
astIoEvent[uiSlot].uliTimeMs := uliIoClockMs;
astIoEvent[uiSlot].usiDirection := usiDirection;
astIoEvent[uiSlot].uiIndex := uiIndex;
astIoEvent[uiSlot].usiKind := usiKind;
astIoEvent[uiSlot].xOld := xOld;
astIoEvent[uiSlot].xNew := xNew;
// Строка кодируется только для изменившегося слота, не для всего FIFO на каждом скане.
sEvent := CONCAT(UDINT_TO_STRING(GVL_HMI.udiIoJournalSequence), ';');
sEvent := CONCAT(sEvent, ULINT_TO_STRING(uliIoClockMs));
sEvent := CONCAT(sEvent, ';'); sEvent := CONCAT(sEvent, USINT_TO_STRING(usiDirection));
sEvent := CONCAT(sEvent, ';'); sEvent := CONCAT(sEvent, UINT_TO_STRING(uiIndex));
sEvent := CONCAT(sEvent, ';'); sEvent := CONCAT(sEvent, USINT_TO_STRING(usiKind));
sEvent := CONCAT(sEvent, ';'); sEvent := CONCAT(sEvent, USINT_TO_STRING(BOOL_TO_USINT(xOld)));
sEvent := CONCAT(sEvent, ';'); sEvent := CONCAT(sEvent, USINT_TO_STRING(BOOL_TO_USINT(xNew)));
GVL_HMI.asIoJournal[uiSlot] := sEvent;
GVL_HMI.uiIoJournalHead := uiSlot;
GVL_HMI.uiIoJournalCount := MIN(UINT#100, GVL_HMI.uiIoJournalCount + UINT#1);
IF NOT xIoSnapshotPublishing THEN
    GVL_HMI.udiIoJournalRevision := GVL_HMI.udiIoJournalRevision + UDINT#1;
END_IF;
END_METHOD

METHOD PRIVATE RunMagazine
auiMagazineEditSlot[1] := GVL_HMI.astMagazineCommand[1].uiEditSlot;
IF auiMagazineEditSlot[1] = UINT#0 THEN
	auiMagazineEditSlot[1] := GVL_HMI.uiMagazineEditSlot;
END_IF;
auiMagazineEditSlot[2] := GVL_HMI.astMagazineCommand[2].uiEditSlot;

fbMagazine1(
	uiMagazineId := UINT#1,
	xInventoryChanged := axMagazineInventoryChanged[1],
	xPointsConfigured := axMagazinePointsReady[1],
	xMechanismReady := (GVL_TWO_PALLET.uiMode = 0) OR GVL_TWO_PALLET.astStatus[1].xReady,
	xTestInitialize := xTestInitializePulse OR xTestAbortActive,
	xTestEnabled := GVL_HMI.stTestScenario.axMagazineEnabled[1],
	stRobotStatus := GVL_ROBOT.Status,
	astMachineStatus := GVL_MACHINE.Status,
	auiMachineType := GVL_MULTI_TYPE.Config.auiMachineType,
	stMagazineCommand := GVL_MAGAZINE.astAutoCommand[1],
	stHmiCommand := GVL_HMI.stRobotCommand,
	xManual := GVL_CELL_CONTROL.xManual AND NOT GVL_CELL_MANAGER.Status.xRunning,
	xIoManual := xIoManualActive,
	xReset := GVL_CELL_CONTROL.xReset OR GVL_HMI.astMagazineCommand[1].xReset OR ((GVL_TWO_PALLET.uiMode = 1) AND (GVL_TWO_PALLET.auiCommand[1] = 16) AND GVL_TWO_PALLET.astStatus[1].xCommandAccepted),
	xGlobalError := GVL_CELL_CONTROL.xGlobalError,
	xHmiEnable := ((GVL_TWO_PALLET.uiMode = 0) AND (GVL_HMI.astMagazineCommand[1].xEnable OR GVL_HMI.xMagazineEnable))
		OR ((GVL_TWO_PALLET.uiMode = 1) AND GVL_TWO_PALLET.astStatus[1].xReady
			AND NOT axTwinMagazineExchangeInProgress[1]
			AND NOT fbMagazine1.Status.xEnabled AND NOT fbMagazine1.Status.xFinished),
	xHmiDisable := GVL_HMI.astMagazineCommand[1].xDisable OR GVL_HMI.xMagazineDisable OR ((GVL_TWO_PALLET.uiMode = 1) AND (NOT GVL_TWO_PALLET.astStatus[1].xEnabled OR GVL_TWO_PALLET.astStatus[1].xBusy OR axTwinMagazineExchangeInProgress[1])),
	xHmiFillBlanks := (GVL_TWO_PALLET.uiMode = 0) AND (GVL_HMI.astMagazineCommand[1].xFill OR GVL_HMI.xMagazineFillBlanks),
	xHmiClear := (GVL_TWO_PALLET.uiMode = 0) AND (GVL_HMI.astMagazineCommand[1].xClear OR GVL_HMI.xMagazineClear),
	xHmiCycleSlot := (GVL_TWO_PALLET.uiMode = 0) AND (GVL_HMI.astMagazineCommand[1].xCycleSlot OR GVL_HMI.xMagazineCycleSlot),
	xHmiApplySlot := (GVL_TWO_PALLET.uiMode = 0) AND (GVL_HMI.astMagazineCommand[1].xApplySlot),
	xHmiApplyPitchX := GVL_HMI.astMagazineCommand[1].xApplyPitchX,
	xHmiApplyPitchY := GVL_HMI.astMagazineCommand[1].xApplyPitchY,
	uiHmiEditSlot := auiMagazineEditSlot[1],
	uiHmiEditDetailType := GVL_HMI.astMagazineCommand[1].uiEditDetailType,
	uiHmiEditProductType := GVL_HMI.astMagazineCommand[1].uiEditProductType,
	lrHmiEditPitchX := GVL_HMI.astMagazineCommand[1].lrEditPitchX,
	lrHmiEditPitchY := GVL_HMI.astMagazineCommand[1].lrEditPitchY,
	xRobotOwnsMagazine := (GVL_CELL_MANAGER.Status.uiActiveMagazine = UINT#1)
		AND (GVL_CELL_MANAGER.Status.xRunning OR GVL_ROBOT.Status.xBusy),
	xRobotCanWorkWithMagazine := xRobotInterfaceReady
		AND axMagazinePointsReady[1]
		AND NOT axTwinMagazineExchangeInProgress[1]
		AND NOT GVL_ROBOT.Status.xError,
	xSharedGeometryEditAllowed := NOT GVL_MAGAZINE.astStatus[1].xEnabled
		AND NOT GVL_MAGAZINE.astStatus[2].xEnabled
		AND NOT GVL_HMI.xMagazineEnable
		AND NOT GVL_HMI.astMagazineCommand[1].xEnable
		AND NOT GVL_HMI.astMagazineCommand[2].xEnable,
	uiRows := GVL_CELL_SETTINGS.MagazineRows,
	uiColumns := GVL_CELL_SETTINGS.MagazineColumns,
	uiTypeCount := GVL_MULTI_TYPE.Config.uiTypeCount,
	auiSlotType := GVL_MULTI_TYPE.Config.auiSlotType,
	FaultRequest := astMagazineFaultRequest[1],
	stInventory := GVL_DETAIL.astMagazine[1],
	lrPitchX := GVL_HMI.MagazinePitchX,
	lrPitchY := GVL_HMI.MagazinePitchY,
	Command => GVL_MAGAZINE.astCommand[1],
	Status => GVL_MAGAZINE.astPartStatus[1],
	Diag => GVL_MAGAZINE.astDiag[1],
	Error => GVL_MAGAZINE.astError[1]
);

fbMagazine2(
	uiMagazineId := UINT#2,
	xInventoryChanged := axMagazineInventoryChanged[2],
	xPointsConfigured := axMagazinePointsReady[2],
	xMechanismReady := (GVL_TWO_PALLET.uiMode = 0) OR GVL_TWO_PALLET.astStatus[2].xReady,
	xTestInitialize := xTestInitializePulse OR xTestAbortActive,
	xTestEnabled := GVL_HMI.stTestScenario.axMagazineEnabled[2],
	stRobotStatus := GVL_ROBOT.Status,
	astMachineStatus := GVL_MACHINE.Status,
	auiMachineType := GVL_MULTI_TYPE.Config.auiMachineType,
	stMagazineCommand := GVL_MAGAZINE.astAutoCommand[2],
	stHmiCommand := GVL_HMI.stRobotCommand,
	xManual := GVL_CELL_CONTROL.xManual AND NOT GVL_CELL_MANAGER.Status.xRunning,
	xIoManual := xIoManualActive,
	xReset := GVL_CELL_CONTROL.xReset OR GVL_HMI.astMagazineCommand[2].xReset OR ((GVL_TWO_PALLET.uiMode = 1) AND (GVL_TWO_PALLET.auiCommand[2] = 16) AND GVL_TWO_PALLET.astStatus[2].xCommandAccepted),
	xGlobalError := GVL_CELL_CONTROL.xGlobalError,
	xHmiEnable := ((GVL_TWO_PALLET.uiMode = 0) AND (GVL_HMI.astMagazineCommand[2].xEnable))
		OR ((GVL_TWO_PALLET.uiMode = 1) AND GVL_TWO_PALLET.astStatus[2].xReady
			AND NOT axTwinMagazineExchangeInProgress[2]
			AND NOT fbMagazine2.Status.xEnabled AND NOT fbMagazine2.Status.xFinished),
	xHmiDisable := GVL_HMI.astMagazineCommand[2].xDisable OR ((GVL_TWO_PALLET.uiMode = 1) AND (NOT GVL_TWO_PALLET.astStatus[2].xEnabled OR GVL_TWO_PALLET.astStatus[2].xBusy OR axTwinMagazineExchangeInProgress[2])),
	xHmiFillBlanks := (GVL_TWO_PALLET.uiMode = 0) AND (GVL_HMI.astMagazineCommand[2].xFill),
	xHmiClear := (GVL_TWO_PALLET.uiMode = 0) AND (GVL_HMI.astMagazineCommand[2].xClear),
	xHmiCycleSlot := (GVL_TWO_PALLET.uiMode = 0) AND (GVL_HMI.astMagazineCommand[2].xCycleSlot),
	xHmiApplySlot := (GVL_TWO_PALLET.uiMode = 0) AND (GVL_HMI.astMagazineCommand[2].xApplySlot),
	xHmiApplyPitchX := GVL_HMI.astMagazineCommand[2].xApplyPitchX,
	xHmiApplyPitchY := GVL_HMI.astMagazineCommand[2].xApplyPitchY,
	uiHmiEditSlot := auiMagazineEditSlot[2],
	uiHmiEditDetailType := GVL_HMI.astMagazineCommand[2].uiEditDetailType,
	uiHmiEditProductType := GVL_HMI.astMagazineCommand[2].uiEditProductType,
	lrHmiEditPitchX := GVL_HMI.astMagazineCommand[2].lrEditPitchX,
	lrHmiEditPitchY := GVL_HMI.astMagazineCommand[2].lrEditPitchY,
	xRobotOwnsMagazine := (GVL_CELL_MANAGER.Status.uiActiveMagazine = UINT#2)
		AND (GVL_CELL_MANAGER.Status.xRunning OR GVL_ROBOT.Status.xBusy),
	xRobotCanWorkWithMagazine := xRobotInterfaceReady
		AND axMagazinePointsReady[2]
		AND NOT axTwinMagazineExchangeInProgress[2]
		AND NOT GVL_ROBOT.Status.xError,
	xSharedGeometryEditAllowed := NOT GVL_MAGAZINE.astStatus[1].xEnabled
		AND NOT GVL_MAGAZINE.astStatus[2].xEnabled
		AND NOT GVL_HMI.xMagazineEnable
		AND NOT GVL_HMI.astMagazineCommand[1].xEnable
		AND NOT GVL_HMI.astMagazineCommand[2].xEnable,
	uiRows := GVL_CELL_SETTINGS.MagazineRows,
	uiColumns := GVL_CELL_SETTINGS.MagazineColumns,
	uiTypeCount := GVL_MULTI_TYPE.Config.uiTypeCount,
	auiSlotType := GVL_MULTI_TYPE.Config.auiSlotType,
	FaultRequest := astMagazineFaultRequest[2],
	stInventory := GVL_DETAIL.astMagazine[2],
	lrPitchX := GVL_HMI.MagazinePitchX,
	lrPitchY := GVL_HMI.MagazinePitchY,
	Command => GVL_MAGAZINE.astCommand[2],
	Status => GVL_MAGAZINE.astPartStatus[2],
	Diag => GVL_MAGAZINE.astDiag[2],
	Error => GVL_MAGAZINE.astError[2]
);

// Сохранить физический инвентарь текущей палеты после подтверждённых действий робота.
FOR uiTwin := 1 TO 2 DO
	GVL_MAGAZINE.astStatus[uiTwin] := GVL_MAGAZINE.astPartStatus[uiTwin];
	IF NOT GVL_TWO_PALLET.astStatus[uiTwin].xError THEN axTwinRobotStopLatched[uiTwin] := FALSE;
	ELSIF GVL_ROBOT.Status.uiMagazineContext = uiTwin THEN axTwinRobotStopLatched[uiTwin] := TRUE; END_IF;
	IF GVL_TWO_PALLET.uiMode = 1 THEN
		uiTwinPallet := GVL_TWO_PALLET.astStatus[uiTwin].uiRobotPallet;
		IF (uiTwinPallet >= UINT#1) AND (uiTwinPallet <= UINT#2) THEN
			GVL_TWO_PALLET.astStore[uiTwin].astPallet[uiTwinPallet] := GVL_DETAIL.astMagazine[uiTwin];
		END_IF;
		GVL_MAGAZINE.astStatus[uiTwin].xReady := GVL_MAGAZINE.astStatus[uiTwin].xReady AND GVL_TWO_PALLET.astStatus[uiTwin].xReady;
		GVL_MAGAZINE.astStatus[uiTwin].xEnableSequenceAllowed := GVL_TWO_PALLET.astStatus[uiTwin].xEnableAllowed;
		GVL_MAGAZINE.astStatus[uiTwin].xEnabled := GVL_TWO_PALLET.astStatus[uiTwin].xEnabled;
		GVL_MAGAZINE.astStatus[uiTwin].xBusy := GVL_MAGAZINE.astPartStatus[uiTwin].xBusy OR GVL_TWO_PALLET.astStatus[uiTwin].xBusy;
		GVL_MAGAZINE.astStatus[uiTwin].xFillAllowed := FALSE;
		GVL_MAGAZINE.astStatus[uiTwin].xClearAllowed := FALSE;
		GVL_MAGAZINE.astStatus[uiTwin].xEditAllowed := FALSE;
		GVL_MAGAZINE.astStatus[uiTwin].xError := GVL_MAGAZINE.astStatus[uiTwin].xError OR GVL_TWO_PALLET.astStatus[uiTwin].xError;
		GVL_MAGAZINE.astError[uiTwin].dwErrorActive := GVL_MAGAZINE.astError[uiTwin].dwErrorActive
			OR GVL_TWO_PALLET.astError[uiTwin].dwErrorActive;
		GVL_MAGAZINE.astError[uiTwin].dwAlarmActive := GVL_MAGAZINE.astError[uiTwin].dwAlarmActive
			OR GVL_TWO_PALLET.astError[uiTwin].dwAlarmActive;
		GVL_MAGAZINE.astStatus[uiTwin].xRobotStopRequired := GVL_MAGAZINE.astStatus[uiTwin].xRobotStopRequired
			OR axTwinRobotStopLatched[uiTwin];
		IF axTwinRobotStopLatched[uiTwin] THEN
			GVL_MAGAZINE.astCommand[uiTwin].xStop := TRUE;
			GVL_MAGAZINE.astCommand[uiTwin].xExecute := FALSE;
		END_IF;
	ELSE
		GVL_TWO_PALLET.astStatic[uiTwin] := GVL_DETAIL.astMagazine[uiTwin];
	END_IF;
END_FOR;

IF GVL_TWO_PALLET.uiMode = 0 THEN
	GVL_TWO_PALLET.lrStaticPitchX := GVL_HMI.MagazinePitchX;
	GVL_TWO_PALLET.lrStaticPitchY := GVL_HMI.MagazinePitchY;
ELSE
	GVL_TWO_PALLET.lrTwinPitchX := GVL_HMI.MagazinePitchX;
	GVL_TWO_PALLET.lrTwinPitchY := GVL_HMI.MagazinePitchY;
END_IF;
END_METHOD

METHOD PRIVATE RunTwoPalletAxis
// Magazine_1/2 — точки привязки Motion: в NORMAL настроить реальные оси EtherCAT.
// MC_Home запускает поиск дома в серводрайвере; FB_AXIS ждёт его Done.
// Ссылки назначаются каждый скан до проверки __ISVALIDREF и вызова FB_AXIS.
GVL_TWO_PALLET.Axis1 REF= Magazine_1;
GVL_TWO_PALLET.Axis2 REF= Magazine_2;
GVL_TWO_PALLET.astInput[1].xAxisBound := __ISVALIDREF(GVL_TWO_PALLET.Axis1);
GVL_TWO_PALLET.astInput[2].xAxisBound := __ISVALIDREF(GVL_TWO_PALLET.Axis2);
FOR uiTwin := 1 TO 2 DO
	GVL_TWO_PALLET.astAxis[uiTwin].Command.xEnable := GVL_TWO_PALLET.astOutput[uiTwin].xPowerOn;
	GVL_TWO_PALLET.astAxis[uiTwin].Command.xDisable := GVL_TWO_PALLET.astOutput[uiTwin].xPowerOff
		OR (GVL_TWO_PALLET.uiMode = 0);
	GVL_TWO_PALLET.astAxis[uiTwin].Command.xPowerPermit := (GVL_TWO_PALLET.uiMode = 1)
		AND CELL_SAFETY.Status.xReady AND GVL_TWO_PALLET.astInput[uiTwin].xIoMapped;
	GVL_TWO_PALLET.astAxis[uiTwin].Command.xGlobalError := GVL_CELL_CONTROL.xGlobalError;
	GVL_TWO_PALLET.astAxis[uiTwin].Command.xResetAllError := GVL_TWO_PALLET.astOutput[uiTwin].xDriveReset;
	GVL_TWO_PALLET.astAxis[uiTwin].Command.xStop := GVL_TWO_PALLET.astOutput[uiTwin].xStop OR GVL_HMI.xIoEmergencyStopActive;
	GVL_TWO_PALLET.astAxis[uiTwin].Command.xHome := GVL_TWO_PALLET.astOutput[uiTwin].xHome;
	GVL_TWO_PALLET.astAxis[uiTwin].Command.xMoveAbsolute := GVL_TWO_PALLET.astOutput[uiTwin].xMove;
	GVL_TWO_PALLET.astAxis[uiTwin].Command.xJogPositive := GVL_TWO_PALLET.astOutput[uiTwin].xJogPositive;
	GVL_TWO_PALLET.astAxis[uiTwin].Command.xJogNegative := GVL_TWO_PALLET.astOutput[uiTwin].xJogNegative;
	GVL_TWO_PALLET.astAxis[uiTwin].MotionParam.lrTargetPosition := GVL_TWO_PALLET.astOutput[uiTwin].lrTarget;
	GVL_TWO_PALLET.astAxis[uiTwin].MotionParam.lrHomePosition := GVL_TWO_PALLET.astActiveConfig[uiTwin].lrHome;
	GVL_TWO_PALLET.astAxis[uiTwin].MotionParam.lrVelocity := GVL_TWO_PALLET.astActiveConfig[uiTwin].lrVelocity;
	GVL_TWO_PALLET.astAxis[uiTwin].MotionParam.lrAcceleration := GVL_TWO_PALLET.astActiveConfig[uiTwin].lrAcceleration;
	GVL_TWO_PALLET.astAxis[uiTwin].MotionParam.lrDeceleration := GVL_TWO_PALLET.astActiveConfig[uiTwin].lrDeceleration;
	GVL_TWO_PALLET.astAxis[uiTwin].MotionParam.lrJerk := GVL_TWO_PALLET.astActiveConfig[uiTwin].lrJerk;
	GVL_TWO_PALLET.astAxis[uiTwin].Timeouts := GVL_CELL_SETTINGS.stAxisTimeouts;
	GVL_TWO_PALLET.astAxis[uiTwin].Timeouts.tHomeTimeout := GVL_TWO_PALLET.astActiveConfig[uiTwin].tHome;
	GVL_TWO_PALLET.astAxis[uiTwin].Timeouts.tMoveTimeout := GVL_TWO_PALLET.astActiveConfig[uiTwin].tMove;
END_FOR;
IF __ISVALIDREF(GVL_TWO_PALLET.Axis1) THEN
	TWIN_AXIS_1(Axis := GVL_TWO_PALLET.Axis1, AxisData := GVL_TWO_PALLET.astAxis[1],
		xResetPermit := GVL_CELL_CONTROL.xManual AND NOT GVL_CELL_MANAGER.Status.xRunning);
END_IF;
IF __ISVALIDREF(GVL_TWO_PALLET.Axis2) THEN
	TWIN_AXIS_2(Axis := GVL_TWO_PALLET.Axis2, AxisData := GVL_TWO_PALLET.astAxis[2],
		xResetPermit := GVL_CELL_CONTROL.xManual AND NOT GVL_CELL_MANAGER.Status.xRunning);
END_IF;
FOR uiTwin := 1 TO 2 DO
	GVL_TWO_PALLET.astInput[uiTwin].xPowered := GVL_TWO_PALLET.astAxis[uiTwin].Status.xPowered;
	GVL_TWO_PALLET.astInput[uiTwin].xHomed := GVL_TWO_PALLET.astAxis[uiTwin].Status.xHomed;
	GVL_TWO_PALLET.astInput[uiTwin].xStandstill := GVL_TWO_PALLET.astAxis[uiTwin].Status.xStandstill;
	GVL_TWO_PALLET.astInput[uiTwin].xDriveError := GVL_TWO_PALLET.astAxis[uiTwin].Status.xError;
	GVL_TWO_PALLET.astInput[uiTwin].xMotionDone := GVL_TWO_PALLET.astAxis[uiTwin].Status.xDone;
	GVL_TWO_PALLET.astInput[uiTwin].lrPosition := GVL_TWO_PALLET.astAxis[uiTwin].Status.lrActualPosition;
	TWIN_SIM[uiTwin](
		xEnable := (GVL_TWO_PALLET.uiMode = UINT#1)
			AND (GVL_CELL_SETTINGS.eTestEnvironment = E_CELL_TEST_ENVIRONMENT.SIMULATION),
		uiP1Signals := GVL_TWO_PALLET.astActiveConfig[uiTwin].uiP1Signals,
		Command := GVL_TWO_PALLET.astOutput[uiTwin]);
	IF (GVL_TWO_PALLET.uiMode = UINT#1)
		AND (GVL_CELL_SETTINGS.eTestEnvironment = E_CELL_TEST_ENVIRONMENT.SIMULATION) THEN
		GVL_TWO_PALLET.astInput[uiTwin].xIoMapped := TRUE;
		GVL_TWO_PALLET.astInput[uiTwin].xLiftDown := TWIN_SIM[uiTwin].xLiftDown;
		GVL_TWO_PALLET.astInput[uiTwin].xLiftUp := TWIN_SIM[uiTwin].xLiftUp;
		GVL_TWO_PALLET.astInput[uiTwin].xLockIn := TWIN_SIM[uiTwin].xLockIn;
		GVL_TWO_PALLET.astInput[uiTwin].xLockOut := TWIN_SIM[uiTwin].xLockOut;
		GVL_TWO_PALLET.astInput[uiTwin].xStopIn := TWIN_SIM[uiTwin].xStopIn;
		GVL_TWO_PALLET.astInput[uiTwin].xStopOut := TWIN_SIM[uiTwin].xStopOut;
		GVL_TWO_PALLET.astInput[uiTwin].xLimitNegative := FALSE;
		GVL_TWO_PALLET.astInput[uiTwin].xLimitPositive := FALSE;
		GVL_TWO_PALLET.astInput[uiTwin].xHomeSensor := GVL_TWO_PALLET.astInput[uiTwin].xHomed
			AND (ABS(GVL_TWO_PALLET.astInput[uiTwin].lrPosition
				- GVL_TWO_PALLET.astActiveConfig[uiTwin].lrHome)
				<= GVL_TWO_PALLET.astActiveConfig[uiTwin].lrTolerance);
		axTwinSimIoOwned[uiTwin] := TRUE;
	ELSIF axTwinSimIoOwned[uiTwin]
	AND (GVL_CELL_SETTINGS.eTestEnvironment <> E_CELL_TEST_ENVIRONMENT.NORMAL) THEN
		// После выхода из виртуальной среды не оставляем её герконы как реальные.
		GVL_TWO_PALLET.astInput[uiTwin].xIoMapped := FALSE;
		GVL_TWO_PALLET.astInput[uiTwin].xLiftDown := FALSE;
		GVL_TWO_PALLET.astInput[uiTwin].xLiftUp := FALSE;
		GVL_TWO_PALLET.astInput[uiTwin].xLockIn := FALSE;
		GVL_TWO_PALLET.astInput[uiTwin].xLockOut := FALSE;
		GVL_TWO_PALLET.astInput[uiTwin].xStopIn := FALSE;
		GVL_TWO_PALLET.astInput[uiTwin].xStopOut := FALSE;
		GVL_TWO_PALLET.astInput[uiTwin].xLimitNegative := FALSE;
		GVL_TWO_PALLET.astInput[uiTwin].xLimitPositive := FALSE;
		GVL_TWO_PALLET.astInput[uiTwin].xHomeSensor := FALSE;
		axTwinSimIoOwned[uiTwin] := FALSE;
	END_IF;
	IF GVL_CELL_SETTINGS.eTestEnvironment = E_CELL_TEST_ENVIRONMENT.NORMAL THEN
		// ReadPhysicalInputs уже заменил виртуальные герконы в начале скана.
		// Концевики и датчик дома заведены в драйвер, не в DI ячейки. Эти legacy-
		// поля не имитируют PDO; результат Home приходит выше через xHomed/xMotionDone.
		GVL_TWO_PALLET.astInput[uiTwin].xLimitNegative := FALSE;
		GVL_TWO_PALLET.astInput[uiTwin].xLimitPositive := FALSE;
		GVL_TWO_PALLET.astInput[uiTwin].xHomeSensor := FALSE;
		axTwinSimIoOwned[uiTwin] := FALSE;
	END_IF;
END_FOR;
END_METHOD

METHOD PRIVATE ReadIoEmergencyStop
// Отдельный канал: останов не ждёт текущую транзакцию подмены I/O.
xIoEmergencyResetRequested := FALSE;
xIoEmergencyResetRejected := FALSE;
udiIoEmergencyRequestSeq := GVL_HMI.udiIoEmergencyCommandSeq;
IF xIoInitialized AND (udiIoEmergencyRequestSeq <> GVL_HMI.udiIoEmergencyAckSeq) THEN
    IF GVL_HMI.uiIoEmergencyAction = UINT#1 THEN
        xIoManualActive := FALSE;
        GVL_HMI.xIoEmergencyStopActive := TRUE;
        GVL_HMI.uiIoEmergencyResult := UINT#1;
        GVL_HMI.udiIoEmergencyAckSeq := udiIoEmergencyRequestSeq;
    ELSE
        xIoEmergencyResetRequested := TRUE;
    END_IF;
END_IF;
IF GVL_HMI.xIoEmergencyStopActive THEN
    GVL_CELL_CONTROL.xStop := TRUE;
    GVL_CELL_CONTROL.xStart := FALSE;
    GVL_CELL_CONTROL.xEnable := FALSE;
    GVL_CELL_CONTROL.xManual := TRUE;
    GVL_ROBOT.Command.xExecute := FALSE;
    GVL_ROBOT.Command.xStop := TRUE;
    GVL_ROBOT.ModbusCommand.xExecute := FALSE;
    GVL_ROBOT.ModbusCommand.xStop := TRUE;
    GVL_HMI.xRobotManualExecute := FALSE;
    GVL_HMI.stRobotCommand.xExecute := FALSE;
    xPointCheckStopRequest := xPointCheckActive;
    FOR uiIoIndex := UINT#1 TO UINT#3 DO
        GVL_HMI.astAxisHmiCommand[uiIoIndex].xJogPositive := FALSE;
        GVL_HMI.astAxisHmiCommand[uiIoIndex].xJogNegative := FALSE;
        GVL_HMI.astAxisHmiCommand[uiIoIndex].xHome := FALSE;
        GVL_HMI.astAxisHmiCommand[uiIoIndex].xMoveAbsolute := FALSE;
        GVL_HMI.astAxisHmiCommand[uiIoIndex].xMoveRelative := FALSE;
        GVL_HMI.axMachineManualHatchOpen[uiIoIndex] := FALSE;
        GVL_HMI.axMachineManualHatchClose[uiIoIndex] := FALSE;
        GVL_HMI.axMachineManualHatchUnlock[uiIoIndex] := FALSE;
        GVL_HMI.axMachineManualHatchLock[uiIoIndex] := FALSE;
        GVL_HMI.axMachineManualChuckOpen[uiIoIndex] := FALSE;
        GVL_HMI.axMachineManualChuckClose[uiIoIndex] := FALSE;
    END_FOR;
END_IF;
END_METHOD

METHOD PRIVATE RunMotion
xManualRecoveryActive := GVL_CELL_CONTROL.xGlobalError
	AND GVL_CELL_CONTROL.xManual
	AND NOT GVL_CELL_MANAGER.Status.xRunning
	AND NOT GVL_HMI.xModbusMode
	AND xHmiConnectionAlive;

// В recovery общая ошибка остаётся на уровне ячейки, но не создаёт каскадную
// ошибку исправных осей. Ниже для этого состояния разрешён только Jog.
GVL_AXIS.arrAxis[1].Command.xGlobalError := GVL_CELL_CONTROL.xGlobalError AND NOT xManualRecoveryActive;
GVL_AXIS.arrAxis[2].Command.xGlobalError := GVL_CELL_CONTROL.xGlobalError AND NOT xManualRecoveryActive;
GVL_AXIS.arrAxis[3].Command.xGlobalError := GVL_CELL_CONTROL.xGlobalError AND NOT xManualRecoveryActive;
GVL_AXIS_GROUP.AxisGroup.Command.xGlobalError := GVL_CELL_CONTROL.xGlobalError AND NOT xManualRecoveryActive;

GVL_AXIS.arrAxis[1].Command.xPowerPermit := NOT GVL_AXIS.arrAxis[1].Command.xGlobalError;
GVL_AXIS.arrAxis[2].Command.xPowerPermit := NOT GVL_AXIS.arrAxis[2].Command.xGlobalError;
GVL_AXIS.arrAxis[3].Command.xPowerPermit := NOT GVL_AXIS.arrAxis[3].Command.xGlobalError;
GVL_AXIS_GROUP.AxisGroup.Command.xPowerPermit := NOT GVL_AXIS_GROUP.AxisGroup.Command.xGlobalError;

// Текущие состояния нужны для единого расчёта разрешений силовых команд.
xRobotMotionCommandActive := (GVL_ROBOT.Diag.eState = E_ROBOT_STATE.MOTION)
	OR (GVL_MOTION_MANAGER.stMotionManager.Diag.eState = E_MOTION_MANAGER_STATE.VALIDATE)
	OR (GVL_MOTION_MANAGER.stMotionManager.Diag.eState = E_MOTION_MANAGER_STATE.MOTION_SIM)
	OR (GVL_MOTION_MANAGER.stMotionManager.Diag.eState = E_MOTION_MANAGER_STATE.DONE);
xDrivesPowered := GVL_AXIS.arrAxis[1].Status.xPowered
	AND GVL_AXIS.arrAxis[2].Status.xPowered
	AND GVL_AXIS.arrAxis[3].Status.xPowered;
xAnyDrivePowered := GVL_AXIS.arrAxis[1].Status.xPowerStageOn
	OR GVL_AXIS.arrAxis[1].Status.xDriveStartOn
	OR GVL_AXIS.arrAxis[2].Status.xPowerStageOn
	OR GVL_AXIS.arrAxis[2].Status.xDriveStartOn
	OR GVL_AXIS.arrAxis[3].Status.xPowerStageOn
	OR GVL_AXIS.arrAxis[3].Status.xDriveStartOn;
xDrivesOff := NOT xAnyDrivePowered
	AND (GVL_AXIS_GROUP.AxisGroup.Diag.iStep = E_AXIS_GROUP_STATE.DISABLED);
xPowerTransitionActive :=
	(GVL_AXIS.arrAxis[1].Diag.iStep = E_AXIS_STATE.POWERING)
	OR (GVL_AXIS.arrAxis[1].Diag.iStep = E_AXIS_STATE.POWERING_DOWN)
	OR (GVL_AXIS.arrAxis[2].Diag.iStep = E_AXIS_STATE.POWERING)
	OR (GVL_AXIS.arrAxis[2].Diag.iStep = E_AXIS_STATE.POWERING_DOWN)
	OR (GVL_AXIS.arrAxis[3].Diag.iStep = E_AXIS_STATE.POWERING)
	OR (GVL_AXIS.arrAxis[3].Diag.iStep = E_AXIS_STATE.POWERING_DOWN)
	OR (GVL_AXIS_GROUP.AxisGroup.Diag.iStep = E_AXIS_GROUP_STATE.ENABLING_POWER)
	OR (GVL_AXIS_GROUP.AxisGroup.Diag.iStep = E_AXIS_GROUP_STATE.ENABLING_GROUP)
	OR (GVL_AXIS_GROUP.AxisGroup.Diag.iStep = E_AXIS_GROUP_STATE.DISABLING_GROUP)
	OR (GVL_AXIS_GROUP.AxisGroup.Diag.iStep = E_AXIS_GROUP_STATE.DISABLING_POWER);
xMotionResetBusy := eMotionResetState <> E_MOTION_RESET_STATE.IDLE;
xAxisDriveError := GVL_AXIS.arrAxis[1].Status.xAxisError
	OR GVL_AXIS.arrAxis[1].Status.xLogicalError
	OR GVL_AXIS.arrAxis[2].Status.xAxisError
	OR GVL_AXIS.arrAxis[2].Status.xLogicalError
	OR GVL_AXIS.arrAxis[3].Status.xAxisError
	OR GVL_AXIS.arrAxis[3].Status.xLogicalError;
xGroupError := GVL_AXIS_GROUP.AxisGroup.Status.xLocalError
	OR GVL_AXIS_GROUP.AxisGroup.Status.xLogicalError
	OR GVL_AXIS_GROUP.AxisGroup.Status.xGroupError;
xDriveError := xAxisDriveError OR xGroupError;
xGroupMotionBusy := GVL_AXIS_GROUP.AxisGroup.Command.xMoveDirect
	OR GVL_AXIS_GROUP.AxisGroup.Command.xMoveLinear
	OR (GVL_AXIS_GROUP.AxisGroup.Diag.iStep = E_AXIS_GROUP_STATE.MOVING_DIRECT)
	OR (GVL_AXIS_GROUP.AxisGroup.Diag.iStep = E_AXIS_GROUP_STATE.MOVING_LINEAR)
	OR (GVL_AXIS_GROUP.AxisGroup.Diag.iStep = E_AXIS_GROUP_STATE.EMG_STOP)
	OR (GVL_AXIS_GROUP.AxisGroup.Diag.iStep = E_AXIS_GROUP_STATE.HALT_STOP)
	OR (GVL_AXIS_GROUP.AxisGroup.Diag.iStep = E_AXIS_GROUP_STATE.WAIT_STOP);
xMotionBusy := GVL_AXIS.arrAxis[1].Status.xMotionBusy
	OR GVL_AXIS.arrAxis[2].Status.xMotionBusy
	OR GVL_AXIS.arrAxis[3].Status.xMotionBusy
	OR xGroupMotionBusy;

// Владелец продолжающейся одиночной команды определяется по автомату FB_AXIS,
// а не по кратковременному импульсу HMI.
uiManualAxisOwner := UINT#0;
FOR uiMachine := 1 TO 3 DO
	IF (uiManualAxisOwner = UINT#0)
	AND (GVL_AXIS.arrAxis[uiMachine].Status.xMotionBusy
		OR (GVL_AXIS.arrAxis[uiMachine].Diag.iStep = E_AXIS_STATE.JOGGING)
		OR (GVL_AXIS.arrAxis[uiMachine].Diag.iStep = E_AXIS_STATE.JOG_DECELERATING)
		OR (GVL_AXIS.arrAxis[uiMachine].Diag.iStep = E_AXIS_STATE.HOMING)
		OR (GVL_AXIS.arrAxis[uiMachine].Diag.iStep = E_AXIS_STATE.MOVE_ABSOLUTE)
		OR (GVL_AXIS.arrAxis[uiMachine].Diag.iStep = E_AXIS_STATE.MOVE_RELATIVE)
		OR (GVL_AXIS.arrAxis[uiMachine].Diag.iStep = E_AXIS_STATE.STOPPING)
		OR (GVL_AXIS.arrAxis[uiMachine].Diag.iStep = E_AXIS_STATE.STOP_RELEASE)) THEN
		uiManualAxisOwner := uiMachine;
	END_IF;
END_FOR;
xMotionBusy := xMotionBusy OR (uiManualAxisOwner > UINT#0);

// Отдельный владелец тестовой динамики ничего не пишет напрямую в существующие
// FB_AXIS/FB_AXIS_GROUP. Он выдаёт им штатные Stop/Disable/Enable-запросы и сам
// вызывает только административные SMC_ChangeDynamicLimits для X/Y/Z.
SIMULATION_DYNAMICS(
	xSimulationMode := GVL_CELL_SETTINGS.eTestEnvironment = E_CELL_TEST_ENVIRONMENT.SIMULATION,
	xSoftMotionMode := NOT GVL_HMI.xModbusMode,
	xAccelerationEnabled := GVL_CELL_SETTINGS.xSimulationAccelerationEnable,
	xPrepareTest := xTestInitializePulse,
	uiRequestedFactor := GVL_CELL_SETTINGS.uiSimulationTimeFactor,
	xCellRunning := GVL_CELL_MANAGER.Status.xRunning,
	xRobotBusy := GVL_ROBOT.Status.xBusy,
	xMotionBusy := xMotionBusy,
	xDrivesPowered := xDrivesPowered,
	xDrivesOff := xDrivesOff,
	eGroupState := GVL_AXIS_GROUP.AxisGroup.Diag.iStep,
	tTransactionTimeout := GVL_CELL_SETTINGS.tSimulationDynamicsTimeout,
	AxisX := X,
	AxisY := Y,
	AxisZ := Z
);
GVL_CELL_CONTROL.xStop := GVL_CELL_CONTROL.xStop OR SIMULATION_DYNAMICS.xCellStopRequest;
xRobotHmiPermit := xRobotHmiPermit AND NOT SIMULATION_DYNAMICS.xBusy;
GVL_CELL_SETTINGS.xSimulationAccelerationActive := SIMULATION_DYNAMICS.xAccelerationActive;
GVL_CELL_SETTINGS.uiSimulationTimeFactorApplied := SIMULATION_DYNAMICS.uiAppliedFactor;
GVL_CELL_SETTINGS.xSimulationAccelerationPending := SIMULATION_DYNAMICS.xPending;
GVL_CELL_SETTINGS.xSimulationAccelerationBusy := SIMULATION_DYNAMICS.xBusy;
GVL_CELL_SETTINGS.xSimulationAccelerationError := SIMULATION_DYNAMICS.xError;
GVL_CELL_SETTINGS.udiSimulationAccelerationErrorId := SIMULATION_DYNAMICS.udiErrorId;

rRobotManualEffectiveSpeedPercent := GVL_HMI.rRobotManualSpeedPercent;
IF xMobileMotionLeaseActive THEN
	// Последний рубеж лимита находится в PLC, а не в браузере или gateway.
	rRobotManualEffectiveSpeedPercent := MIN(
		rRobotManualEffectiveSpeedPercent,
		rMobileMotionSpeedLimitPercent
	);
END_IF;

GVL_HMI.stRobotHmiStatus.xDrivesPowered := xDrivesPowered;
GVL_HMI.stRobotHmiStatus.xDrivesOff := xDrivesOff;
GVL_HMI.stRobotHmiStatus.xPowerTransitionActive := xPowerTransitionActive;
GVL_HMI.stRobotHmiStatus.xDrivesEnableAllowed := xRobotHmiPermit
	AND xHmiConnectionAlive
	AND NOT GVL_HMI.xModbusMode
	AND (NOT GVL_CELL_CONTROL.xGlobalError OR xManualRecoveryActive)
	AND xDrivesOff
	AND NOT xAxisDriveError
	AND NOT xRobotMotionCommandActive
	AND NOT xMotionBusy
	AND NOT xMotionResetBusy;
GVL_HMI.stRobotHmiStatus.xDrivesDisableAllowed := xRobotHmiPermit
	AND xHmiConnectionAlive
	AND NOT GVL_HMI.xModbusMode
	AND (xAnyDrivePowered
		OR (GVL_AXIS_GROUP.AxisGroup.Diag.iStep = E_AXIS_GROUP_STATE.READY))
	AND NOT xPowerTransitionActive
	AND NOT xRobotMotionCommandActive
	AND NOT xMotionBusy
	AND NOT xMotionResetBusy;
GVL_HMI.stRobotHmiStatus.xResetAllowed := xRobotHmiPermit
	AND xHmiConnectionAlive
	AND NOT GVL_HMI.xModbusMode
	AND (NOT GVL_CELL_CONTROL.xGlobalError OR xManualRecoveryActive)
	AND NOT xMotionBusy
	AND NOT xMotionResetBusy;
GVL_HMI.stRobotHmiStatus.xStopAllowed := xRobotHmiPermit
	AND xHmiConnectionAlive
	AND NOT GVL_HMI.xModbusMode
	AND (xMotionBusy OR xRobotMotionCommandActive);

// Решение о приёме фиксируется до вызова Motion FB. Позднее фактический статус
// может измениться в том же цикле и не должен превращать принятую команду в отказ.
xHmiDrivesEnableAccepted := GVL_HMI.xRobotDrivesEnable
	AND GVL_HMI.stRobotHmiStatus.xDrivesEnableAllowed;
xHmiDrivesDisableAccepted := GVL_HMI.xRobotDrivesDisable
	AND GVL_HMI.stRobotHmiStatus.xDrivesDisableAllowed;
xHmiResetAccepted := GVL_HMI.xRobotReset
	AND GVL_HMI.stRobotHmiStatus.xResetAllowed;
xHmiStopAccepted := GVL_HMI.xRobotStop
	AND GVL_HMI.stRobotHmiStatus.xStopAllowed;

xMotionResetRequest := NOT GVL_HMI.xModbusMode
	AND (GVL_CELL_CONTROL.xReset OR xHmiResetAccepted);
rtMotionReset(CLK := xMotionResetRequest);
xGroupResetPulse := FALSE;
xAxisResetPulse := FALSE;

// MC_GroupReset самостоятельно сбрасывает все оси группы. Локальные FB_AXIS
// получают отдельный последующий импульс только для очистки своих защёлок.
CASE eMotionResetState OF
	E_MOTION_RESET_STATE.IDLE:
		IF rtMotionReset.Q THEN
			eMotionResetState := E_MOTION_RESET_STATE.RESET_GROUP;
		END_IF;

	E_MOTION_RESET_STATE.RESET_GROUP:
		xGroupResetPulse := TRUE;
		eMotionResetState := E_MOTION_RESET_STATE.WAIT_GROUP;

	E_MOTION_RESET_STATE.WAIT_GROUP:
		IF (GVL_AXIS_GROUP.AxisGroup.Diag.iStep <> E_AXIS_GROUP_STATE.ERROR)
		AND (GVL_AXIS_GROUP.AxisGroup.Diag.iStep <> E_AXIS_GROUP_STATE.RESETTING)
		AND (GVL_AXIS_GROUP.AxisGroup.Diag.iStep <> E_AXIS_GROUP_STATE.RESET_VERIFY)
		AND NOT GVL_AXIS_GROUP.AxisGroup.Status.xLocalError THEN
			eMotionResetState := E_MOTION_RESET_STATE.RESET_AXES;
		ELSIF (GVL_AXIS_GROUP.AxisGroup.Diag.iStep = E_AXIS_GROUP_STATE.ERROR) THEN
			// Один запрос оператора формирует только один импульс. Если активная причина
			// ещё не снялась, следующий reset должен быть отдельной осознанной командой.
			eMotionResetState := E_MOTION_RESET_STATE.IDLE;
		END_IF;

	E_MOTION_RESET_STATE.RESET_AXES:
		xAxisResetPulse := TRUE;
		eMotionResetState := E_MOTION_RESET_STATE.WAIT_AXES;

	E_MOTION_RESET_STATE.WAIT_AXES:
		IF (GVL_AXIS.arrAxis[1].Diag.iStep <> E_AXIS_STATE.RESET_AXIS_ERROR)
		AND (GVL_AXIS.arrAxis[1].Diag.iStep <> E_AXIS_STATE.RESET_RELEASE)
		AND (GVL_AXIS.arrAxis[1].Diag.iStep <> E_AXIS_STATE.RESET_FINISH)
		AND (GVL_AXIS.arrAxis[2].Diag.iStep <> E_AXIS_STATE.RESET_AXIS_ERROR)
		AND (GVL_AXIS.arrAxis[2].Diag.iStep <> E_AXIS_STATE.RESET_RELEASE)
		AND (GVL_AXIS.arrAxis[2].Diag.iStep <> E_AXIS_STATE.RESET_FINISH)
		AND (GVL_AXIS.arrAxis[3].Diag.iStep <> E_AXIS_STATE.RESET_AXIS_ERROR)
		AND (GVL_AXIS.arrAxis[3].Diag.iStep <> E_AXIS_STATE.RESET_RELEASE)
		AND (GVL_AXIS.arrAxis[3].Diag.iStep <> E_AXIS_STATE.RESET_FINISH) THEN
			eMotionResetState := E_MOTION_RESET_STATE.IDLE;
		END_IF;
END_CASE;
xMotionResetBusy := eMotionResetState <> E_MOTION_RESET_STATE.IDLE;

GVL_AXIS.arrAxis[1].Command.xResetAllError := xAxisResetPulse;
GVL_AXIS.arrAxis[2].Command.xResetAllError := xAxisResetPulse;
GVL_AXIS.arrAxis[3].Command.xResetAllError := xAxisResetPulse;
GVL_AXIS_GROUP.AxisGroup.Command.xReset := xGroupResetPulse;

GVL_AXIS.arrAxis[1].Command.xEnable := (GVL_CELL_CONTROL.xEnable
	AND NOT GVL_HMI.xModbusMode
	AND NOT GVL_HMI.xRobotControlModeApply)
	OR xHmiDrivesEnableAccepted
	OR SIMULATION_DYNAMICS.xDrivesEnableRequest;
GVL_AXIS.arrAxis[2].Command.xEnable := (GVL_CELL_CONTROL.xEnable
	AND NOT GVL_HMI.xModbusMode
	AND NOT GVL_HMI.xRobotControlModeApply)
	OR xHmiDrivesEnableAccepted
	OR SIMULATION_DYNAMICS.xDrivesEnableRequest;
GVL_AXIS.arrAxis[3].Command.xEnable := (GVL_CELL_CONTROL.xEnable
	AND NOT GVL_HMI.xModbusMode
	AND NOT GVL_HMI.xRobotControlModeApply)
	OR xHmiDrivesEnableAccepted
	OR SIMULATION_DYNAMICS.xDrivesEnableRequest;
GVL_AXIS_GROUP.AxisGroup.Command.xPowerEnable := (GVL_CELL_CONTROL.xEnable
	AND NOT GVL_HMI.xModbusMode
	AND NOT GVL_HMI.xRobotControlModeApply)
	OR xHmiDrivesEnableAccepted
	OR SIMULATION_DYNAMICS.xDrivesEnableRequest;

xPowerDisableRequest := GVL_CELL_CONTROL.xDisable OR xRobotAutoPowerOff
	OR xHmiDrivesDisableAccepted
	OR SIMULATION_DYNAMICS.xGroupDisableRequest;
GVL_AXIS_GROUP.AxisGroup.Command.xDisable := xPowerDisableRequest;
// Сначала группа обязана перейти в GroupDisabled. Только её OFF_REQUEST
// разрешает FB_AXIS снять DriveStart и RegulatorOn.
GVL_AXIS.arrAxis[1].Command.xDisable :=
	(GVL_AXIS_GROUP.AxisGroup.Diag.iPowerMode = E_AXIS_GROUP_POWER_MODE.OFF_REQUEST)
	OR (xPowerDisableRequest
		AND (GVL_AXIS_GROUP.AxisGroup.Diag.iStep = E_AXIS_GROUP_STATE.DISABLED));
GVL_AXIS.arrAxis[2].Command.xDisable := GVL_AXIS.arrAxis[1].Command.xDisable;
GVL_AXIS.arrAxis[3].Command.xDisable := GVL_AXIS.arrAxis[1].Command.xDisable;

// Stop получает только текущий владелец движения: одна ось либо координатная группа.
GVL_AXIS.arrAxis[1].Command.xStop := ((xHmiStopAccepted AND NOT GVL_HMI.xModbusMode)
	OR xMobileMotionStopRequest
	OR SIMULATION_DYNAMICS.xMotionStopRequest OR xIoManualActive OR GVL_HMI.xIoEmergencyStopActive)
	AND NOT xGroupMotionBusy AND (uiManualAxisOwner = UINT#1);
GVL_AXIS.arrAxis[2].Command.xStop := ((xHmiStopAccepted AND NOT GVL_HMI.xModbusMode)
	OR xMobileMotionStopRequest
	OR SIMULATION_DYNAMICS.xMotionStopRequest OR xIoManualActive OR GVL_HMI.xIoEmergencyStopActive)
	AND NOT xGroupMotionBusy AND (uiManualAxisOwner = UINT#2);
GVL_AXIS.arrAxis[3].Command.xStop := ((xHmiStopAccepted AND NOT GVL_HMI.xModbusMode)
	OR xMobileMotionStopRequest
	OR SIMULATION_DYNAMICS.xMotionStopRequest OR xIoManualActive OR GVL_HMI.xIoEmergencyStopActive)
	AND NOT xGroupMotionBusy AND (uiManualAxisOwner = UINT#3);
GVL_AXIS_GROUP.AxisGroup.Command.xStopCmd :=
	NOT GVL_HMI.xModbusMode
	AND (xHmiStopAccepted OR xRobotProgramStopRequest OR xPointCheckStopRequest
		OR xPointCheckStopping OR SIMULATION_DYNAMICS.xMotionStopRequest OR xIoManualActive OR GVL_HMI.xIoEmergencyStopActive)
	AND xGroupMotionBusy;

// Из новых запросов также выбирается только одна ось. Если движение уже идёт,
// запрос другой оси будет отклонён ниже без передачи в FB_AXIS.
uiManualAxisRequest := UINT#0;
FOR uiMachine := 1 TO 3 DO
	artHmiAxisHome[uiMachine](CLK := GVL_HMI.astAxisHmiCommand[uiMachine].xHome);
	artHmiAxisMoveAbsolute[uiMachine](CLK := GVL_HMI.astAxisHmiCommand[uiMachine].xMoveAbsolute);
	artHmiAxisMoveRelative[uiMachine](CLK := GVL_HMI.astAxisHmiCommand[uiMachine].xMoveRelative);
	axHmiAxisHomePulse[uiMachine] := artHmiAxisHome[uiMachine].Q;
	axHmiAxisMoveAbsolutePulse[uiMachine] := artHmiAxisMoveAbsolute[uiMachine].Q;
	axHmiAxisMoveRelativePulse[uiMachine] := artHmiAxisMoveRelative[uiMachine].Q;

	IF (GVL_HMI.astAxisHmiCommand[uiMachine].xJogPositive
		OR GVL_HMI.astAxisHmiCommand[uiMachine].xJogNegative
		OR axHmiAxisHomePulse[uiMachine]
		OR axHmiAxisMoveAbsolutePulse[uiMachine]
		OR axHmiAxisMoveRelativePulse[uiMachine])
	AND (uiManualAxisRequest = UINT#0) THEN
		uiManualAxisRequest := uiMachine;
	END_IF;
END_FOR;
IF uiManualAxisOwner = UINT#0 THEN
	uiManualAxisOwner := uiManualAxisRequest;
END_IF;

FOR uiMachine := 1 TO 3 DO
	CASE uiMachine OF
		1:
			axRobotSoftwareLimitsEnabled[uiMachine] := X.bSWLimitEnable;
			alrRobotSoftwareMinPosition[uiMachine] := X.fSWLimitNegative;
			alrRobotSoftwareMaxPosition[uiMachine] := X.fSWLimitPositive;
			alrRobotManualRatedVelocity[uiMachine] := X.fSWMaxVelocity;
			IF alrRobotManualRatedVelocity[uiMachine] <= 0.0 THEN
				alrRobotManualRatedVelocity[uiMachine] := X.fMaxVelocity;
			END_IF;
			alrRobotRatedAcceleration[uiMachine] := X.fSWMaxAcceleration;
			IF alrRobotRatedAcceleration[uiMachine] <= 0.0 THEN
				alrRobotRatedAcceleration[uiMachine] := X.fMaxAcceleration;
			END_IF;
			alrRobotRatedDeceleration[uiMachine] := X.fSWMaxDeceleration;
			IF alrRobotRatedDeceleration[uiMachine] <= 0.0 THEN
				alrRobotRatedDeceleration[uiMachine] := X.fMaxDeceleration;
			END_IF;
			alrRobotRatedJerk[uiMachine] := X.fSWMaxJerk;
			IF alrRobotRatedJerk[uiMachine] <= 0.0 THEN
				alrRobotRatedJerk[uiMachine] := X.fMaxJerk;
			END_IF;
		2:
			axRobotSoftwareLimitsEnabled[uiMachine] := Y.bSWLimitEnable;
			alrRobotSoftwareMinPosition[uiMachine] := Y.fSWLimitNegative;
			alrRobotSoftwareMaxPosition[uiMachine] := Y.fSWLimitPositive;
			alrRobotManualRatedVelocity[uiMachine] := Y.fSWMaxVelocity;
			IF alrRobotManualRatedVelocity[uiMachine] <= 0.0 THEN
				alrRobotManualRatedVelocity[uiMachine] := Y.fMaxVelocity;
			END_IF;
			alrRobotRatedAcceleration[uiMachine] := Y.fSWMaxAcceleration;
			IF alrRobotRatedAcceleration[uiMachine] <= 0.0 THEN
				alrRobotRatedAcceleration[uiMachine] := Y.fMaxAcceleration;
			END_IF;
			alrRobotRatedDeceleration[uiMachine] := Y.fSWMaxDeceleration;
			IF alrRobotRatedDeceleration[uiMachine] <= 0.0 THEN
				alrRobotRatedDeceleration[uiMachine] := Y.fMaxDeceleration;
			END_IF;
			alrRobotRatedJerk[uiMachine] := Y.fSWMaxJerk;
			IF alrRobotRatedJerk[uiMachine] <= 0.0 THEN
				alrRobotRatedJerk[uiMachine] := Y.fMaxJerk;
			END_IF;
		3:
			axRobotSoftwareLimitsEnabled[uiMachine] := Z.bSWLimitEnable;
			alrRobotSoftwareMinPosition[uiMachine] := Z.fSWLimitNegative;
			alrRobotSoftwareMaxPosition[uiMachine] := Z.fSWLimitPositive;
			alrRobotManualRatedVelocity[uiMachine] := Z.fSWMaxVelocity;
			IF alrRobotManualRatedVelocity[uiMachine] <= 0.0 THEN
				alrRobotManualRatedVelocity[uiMachine] := Z.fMaxVelocity;
			END_IF;
			alrRobotRatedAcceleration[uiMachine] := Z.fSWMaxAcceleration;
			IF alrRobotRatedAcceleration[uiMachine] <= 0.0 THEN
				alrRobotRatedAcceleration[uiMachine] := Z.fMaxAcceleration;
			END_IF;
			alrRobotRatedDeceleration[uiMachine] := Z.fSWMaxDeceleration;
			IF alrRobotRatedDeceleration[uiMachine] <= 0.0 THEN
				alrRobotRatedDeceleration[uiMachine] := Z.fMaxDeceleration;
			END_IF;
			alrRobotRatedJerk[uiMachine] := Z.fSWMaxJerk;
			IF alrRobotRatedJerk[uiMachine] <= 0.0 THEN
				alrRobotRatedJerk[uiMachine] := Z.fMaxJerk;
			END_IF;
	END_CASE;
	IF alrRobotManualRatedVelocity[uiMachine] <= 0.0 THEN
		alrRobotManualRatedVelocity[uiMachine] := alrRobotManualFallbackVelocity[uiMachine];
	END_IF;
	IF alrRobotRatedAcceleration[uiMachine] <= 0.0 THEN
		alrRobotRatedAcceleration[uiMachine] := alrRobotManualAcceleration[uiMachine];
	END_IF;
	IF alrRobotRatedDeceleration[uiMachine] <= 0.0 THEN
		alrRobotRatedDeceleration[uiMachine] := alrRobotManualDeceleration[uiMachine];
	END_IF;
	IF alrRobotRatedJerk[uiMachine] <= 0.0 THEN
		alrRobotRatedJerk[uiMachine] := alrRobotManualJerk[uiMachine];
	END_IF;
	axRobotSoftwareLimitsEnabled[uiMachine] := axRobotSoftwareLimitsEnabled[uiMachine]
		AND (alrRobotSoftwareMaxPosition[uiMachine] > alrRobotSoftwareMinPosition[uiMachine]);
	GVL_HMI.astAxisHmiStatus[uiMachine].lrMinPosition := alrRobotSoftwareMinPosition[uiMachine];
	GVL_HMI.astAxisHmiStatus[uiMachine].lrMaxPosition := alrRobotSoftwareMaxPosition[uiMachine];
	// Для JOG и одиночных перемещений коэффициент применяется непосредственно
	// к входу Velocity соответствующего Motion FB.
	alrRobotJogVelocity[uiMachine] := alrRobotManualRatedVelocity[uiMachine]
		* REAL_TO_LREAL(rRobotManualEffectiveSpeedPercent) / 100.0;

	GVL_AXIS.arrAxis[uiMachine].Command.xJogPositive := FALSE;
	GVL_AXIS.arrAxis[uiMachine].Command.xJogNegative := FALSE;
	GVL_AXIS.arrAxis[uiMachine].Command.xHome := FALSE;
	GVL_AXIS.arrAxis[uiMachine].Command.xMoveAbsolute := FALSE;
	GVL_AXIS.arrAxis[uiMachine].Command.xMoveRelative := FALSE;
	axManualAxisCommandRejected[uiMachine] := FALSE;

	GVL_AXIS.arrAxis[uiMachine].MotionParam.lrVelocity := alrRobotJogVelocity[uiMachine];
	GVL_AXIS.arrAxis[uiMachine].MotionParam.lrAcceleration := alrRobotRatedAcceleration[uiMachine]
		* REAL_TO_LREAL(GVL_CELL_SETTINGS.rRobotAccelerationPercent) / 100.0;
	GVL_AXIS.arrAxis[uiMachine].MotionParam.lrDeceleration := alrRobotRatedDeceleration[uiMachine]
		* REAL_TO_LREAL(GVL_CELL_SETTINGS.rRobotDecelerationPercent) / 100.0;
	GVL_AXIS.arrAxis[uiMachine].MotionParam.lrJerk := alrRobotRatedJerk[uiMachine]
		* REAL_TO_LREAL(GVL_CELL_SETTINGS.rRobotJerkPercent) / 100.0;

	axManualAxisBaseAllowed[uiMachine] := xRobotHmiPermit
		AND NOT GVL_TWO_PALLET.astStatus[1].xBusy AND NOT GVL_TWO_PALLET.astStatus[2].xBusy
		AND NOT xPointCheckActive
		AND xHmiConnectionAlive
		AND NOT GVL_HMI.xModbusMode
		AND (NOT GVL_CELL_CONTROL.xGlobalError OR xManualRecoveryActive)
		AND NOT xDriveError
		AND NOT GVL_ROBOT.Status.xBusy
		AND (GVL_AXIS_GROUP.AxisGroup.Diag.iStep = E_AXIS_GROUP_STATE.READY)
		AND (NOT xMotionBusy OR (uiManualAxisOwner = uiMachine))
		AND GVL_AXIS.arrAxis[uiMachine].Status.xPowered
		AND NOT GVL_AXIS.arrAxis[uiMachine].Status.xAxisError
		AND NOT GVL_AXIS.arrAxis[uiMachine].Status.xLogicalError
		AND (
			((GVL_AXIS.arrAxis[uiMachine].Diag.iStep = E_AXIS_STATE.READY)
				AND GVL_AXIS.arrAxis[uiMachine].Status.xCanStartMotion)
			OR ((uiManualAxisOwner = uiMachine)
				AND ((GVL_AXIS.arrAxis[uiMachine].Diag.iStep = E_AXIS_STATE.JOGGING)
					OR (GVL_AXIS.arrAxis[uiMachine].Diag.iStep = E_AXIS_STATE.JOG_DECELERATING)))
		);
END_FOR;

// Единственный источник допустимого диапазона координат — активные Software Limits
// соответствующих AXIS_REF_SM3. RunMotion выполняется раньше RunRobot, поэтому
// FB_POINT_MANAGER получает актуальный снимок границ до проверки новой точки.
GVL_POINT_MANAGER.PointManager.Diag.lrX_MinLimit := alrRobotSoftwareMinPosition[1];
GVL_POINT_MANAGER.PointManager.Diag.lrX_MaxLimit := alrRobotSoftwareMaxPosition[1];
GVL_POINT_MANAGER.PointManager.Diag.lrY_MinLimit := alrRobotSoftwareMinPosition[2];
GVL_POINT_MANAGER.PointManager.Diag.lrY_MaxLimit := alrRobotSoftwareMaxPosition[2];
GVL_POINT_MANAGER.PointManager.Diag.lrZ_MinLimit := alrRobotSoftwareMinPosition[3];
GVL_POINT_MANAGER.PointManager.Diag.lrZ_MaxLimit := alrRobotSoftwareMaxPosition[3];
GVL_POINT_MANAGER.PointManager.Diag.xXLimitValid := axRobotSoftwareLimitsEnabled[1];
GVL_POINT_MANAGER.PointManager.Diag.xYLimitValid := axRobotSoftwareLimitsEnabled[2];
GVL_POINT_MANAGER.PointManager.Diag.xZLimitValid := axRobotSoftwareLimitsEnabled[3];

IF uiManualAxisRequest > UINT#0 THEN
	FOR uiMachine := 1 TO 3 DO
		IF uiMachine <> uiManualAxisRequest
		AND (GVL_HMI.astAxisHmiCommand[uiMachine].xJogPositive
			OR GVL_HMI.astAxisHmiCommand[uiMachine].xJogNegative
			OR axHmiAxisHomePulse[uiMachine]
			OR axHmiAxisMoveAbsolutePulse[uiMachine]
			OR axHmiAxisMoveRelativePulse[uiMachine]) THEN
			axManualAxisCommandRejected[uiMachine] := TRUE;
		END_IF;
	END_FOR;

	IF uiManualAxisOwner <> uiManualAxisRequest THEN
		axManualAxisCommandRejected[uiManualAxisRequest] := TRUE;
	ELSIF NOT axManualAxisBaseAllowed[uiManualAxisRequest] THEN
		axManualAxisCommandRejected[uiManualAxisRequest] := TRUE;
	ELSIF axHmiAxisHomePulse[uiManualAxisRequest] THEN
		IF NOT GVL_HMI.astAxisHmiCommand[uiManualAxisRequest].xJogPositive
		AND NOT GVL_HMI.astAxisHmiCommand[uiManualAxisRequest].xJogNegative
		AND NOT GVL_HMI.astAxisHmiCommand[uiManualAxisRequest].xMoveAbsolute
		AND NOT GVL_HMI.astAxisHmiCommand[uiManualAxisRequest].xMoveRelative
		AND NOT GVL_CELL_CONTROL.xGlobalError
		AND GVL_AXIS.arrAxis[uiManualAxisRequest].Status.xCanStartMotion THEN
			GVL_AXIS.arrAxis[uiManualAxisRequest].Command.xHome := TRUE;
		ELSE
			axManualAxisCommandRejected[uiManualAxisRequest] := TRUE;
		END_IF;
	ELSIF axHmiAxisMoveAbsolutePulse[uiManualAxisRequest] THEN
		IF NOT GVL_HMI.astAxisHmiCommand[uiManualAxisRequest].xMoveRelative
		AND NOT GVL_HMI.astAxisHmiCommand[uiManualAxisRequest].xJogPositive
		AND NOT GVL_HMI.astAxisHmiCommand[uiManualAxisRequest].xJogNegative
		AND NOT GVL_CELL_CONTROL.xGlobalError
		AND GVL_AXIS.arrAxis[uiManualAxisRequest].Status.xCanStartMotion
		AND (GVL_HMI.astAxisHmiCommand[uiManualAxisRequest].lrTargetPosition
			>= GVL_HMI.astAxisHmiStatus[uiManualAxisRequest].lrMinPosition)
		AND (GVL_HMI.astAxisHmiCommand[uiManualAxisRequest].lrTargetPosition
			<= GVL_HMI.astAxisHmiStatus[uiManualAxisRequest].lrMaxPosition)
		AND (NOT axRobotSoftwareLimitsEnabled[uiManualAxisRequest]
			OR (GVL_HMI.astAxisHmiCommand[uiManualAxisRequest].lrTargetPosition
				>= alrRobotSoftwareMinPosition[uiManualAxisRequest]))
		AND (NOT axRobotSoftwareLimitsEnabled[uiManualAxisRequest]
			OR (GVL_HMI.astAxisHmiCommand[uiManualAxisRequest].lrTargetPosition
				<= alrRobotSoftwareMaxPosition[uiManualAxisRequest])) THEN
			GVL_AXIS.arrAxis[uiManualAxisRequest].MotionParam.lrTargetPosition :=
				GVL_HMI.astAxisHmiCommand[uiManualAxisRequest].lrTargetPosition;
			GVL_AXIS.arrAxis[uiManualAxisRequest].Command.xMoveAbsolute := TRUE;
		ELSE
			axManualAxisCommandRejected[uiManualAxisRequest] := TRUE;
		END_IF;
	ELSIF GVL_HMI.xRobotContinuousMode THEN
		IF (GVL_HMI.astAxisHmiCommand[uiManualAxisRequest].xJogPositive
			XOR GVL_HMI.astAxisHmiCommand[uiManualAxisRequest].xJogNegative)
		AND NOT GVL_HMI.astAxisHmiCommand[uiManualAxisRequest].xMoveAbsolute
		AND NOT GVL_HMI.astAxisHmiCommand[uiManualAxisRequest].xMoveRelative THEN
			IF GVL_HMI.astAxisHmiCommand[uiManualAxisRequest].xJogPositive THEN
				// Направление не снимается упреждающе: software limit контролирует SoftMotion.
				GVL_AXIS.arrAxis[uiManualAxisRequest].Command.xJogPositive := TRUE;
			ELSE
				GVL_AXIS.arrAxis[uiManualAxisRequest].Command.xJogNegative := TRUE;
			END_IF;
		ELSE
			axManualAxisCommandRejected[uiManualAxisRequest] := TRUE;
		END_IF;
	ELSE
		IF axHmiAxisMoveRelativePulse[uiManualAxisRequest]
		AND NOT GVL_HMI.astAxisHmiCommand[uiManualAxisRequest].xMoveAbsolute
		AND NOT GVL_HMI.astAxisHmiCommand[uiManualAxisRequest].xJogPositive
		AND NOT GVL_HMI.astAxisHmiCommand[uiManualAxisRequest].xJogNegative
		AND NOT GVL_CELL_CONTROL.xGlobalError
		AND GVL_AXIS.arrAxis[uiManualAxisRequest].Status.xHomed
		AND GVL_AXIS.arrAxis[uiManualAxisRequest].Status.xCanStartMotion
		AND (ABS(ABS(GVL_HMI.astAxisHmiCommand[uiManualAxisRequest].lrRelativeDistance)
			- GVL_HMI.lrRobotManualStep) < 0.0001)
		AND (GVL_AXIS.arrAxis[uiManualAxisRequest].Status.lrActualPosition
			+ GVL_HMI.astAxisHmiCommand[uiManualAxisRequest].lrRelativeDistance
			>= GVL_HMI.astAxisHmiStatus[uiManualAxisRequest].lrMinPosition)
		AND (GVL_AXIS.arrAxis[uiManualAxisRequest].Status.lrActualPosition
			+ GVL_HMI.astAxisHmiCommand[uiManualAxisRequest].lrRelativeDistance
			<= GVL_HMI.astAxisHmiStatus[uiManualAxisRequest].lrMaxPosition)
		AND (NOT axRobotSoftwareLimitsEnabled[uiManualAxisRequest]
			OR (GVL_AXIS.arrAxis[uiManualAxisRequest].Status.lrActualPosition
				+ GVL_HMI.astAxisHmiCommand[uiManualAxisRequest].lrRelativeDistance
				>= alrRobotSoftwareMinPosition[uiManualAxisRequest]))
		AND (NOT axRobotSoftwareLimitsEnabled[uiManualAxisRequest]
			OR (GVL_AXIS.arrAxis[uiManualAxisRequest].Status.lrActualPosition
				+ GVL_HMI.astAxisHmiCommand[uiManualAxisRequest].lrRelativeDistance
				<= alrRobotSoftwareMaxPosition[uiManualAxisRequest])) THEN
			GVL_AXIS.arrAxis[uiManualAxisRequest].MotionParam.lrDistance :=
				GVL_HMI.astAxisHmiCommand[uiManualAxisRequest].lrRelativeDistance;
			GVL_AXIS.arrAxis[uiManualAxisRequest].Command.xMoveRelative := TRUE;
		ELSE
			axManualAxisCommandRejected[uiManualAxisRequest] := TRUE;
		END_IF;
	END_IF;
END_IF;

// Предупреждение формируется только на фронт действительно отклонённой попытки.
FOR uiMachine := 1 TO 3 DO
	artManualAxisReject[uiMachine](CLK := axManualAxisCommandRejected[uiMachine]);
END_FOR;

// Все оси используют единый инженерный профиль. Настройки принимаются только
// вне переходов питания и движения, поэтому активный шаг не меняет PT на лету.
FOR uiMachine := 1 TO 3 DO
	GVL_AXIS.arrAxis[uiMachine].Timeouts := GVL_CELL_SETTINGS.stAxisTimeouts;
END_FOR;
GVL_AXIS_GROUP.AxisGroup.Timeouts := GVL_CELL_SETTINGS.stAxisGroupTimeouts;

AXIS_X(
	FaultRequest := astAxisFaultRequest[1],
	xResetPermit := xRobotHmiPermit,
	Axis := X,
	AxisData := GVL_AXIS.arrAxis[1]
);
AXIS_Y(
	FaultRequest := astAxisFaultRequest[2],
	xResetPermit := xRobotHmiPermit,
	Axis := Y,
	AxisData := GVL_AXIS.arrAxis[2]
);
AXIS_Z(
	FaultRequest := astAxisFaultRequest[3],
	xResetPermit := xRobotHmiPermit,
	Axis := Z,
	AxisData := GVL_AXIS.arrAxis[3]
);

FOR uiMachine := 1 TO 3 DO
	IF artManualAxisReject[uiMachine].Q THEN
		GVL_AXIS.arrAxis[uiMachine].Diag.stWarning.uiCode := WRN_HMI_MANUAL_REJECTED;
		GVL_AXIS.arrAxis[uiMachine].Diag.stWarning.udiSequence :=
			GVL_AXIS.arrAxis[uiMachine].Diag.stWarning.udiSequence + UDINT#1;
		IF GVL_AXIS.arrAxis[uiMachine].Diag.stWarning.udiSequence = UDINT#0 THEN
			GVL_AXIS.arrAxis[uiMachine].Diag.stWarning.udiSequence := UDINT#1;
		END_IF;
	END_IF;
END_FOR;

// Запрошенный коэффициент живёт отдельно от применённого. Таймеры моделей и
// динамика осей получают только значение, подтверждённое отдельным FB на границе теста.
IF GVL_CELL_SETTINGS.uiSimulationTimeFactor < UINT#1 THEN
	GVL_CELL_SETTINGS.uiSimulationTimeFactor := UINT#1;
ELSIF GVL_ROBOT_MODBUS.xModeActive
AND (GVL_CELL_SETTINGS.uiSimulationTimeFactor > UINT#250) THEN
	GVL_CELL_SETTINGS.uiSimulationTimeFactor := UINT#250;
ELSIF NOT GVL_ROBOT_MODBUS.xModeActive
AND (GVL_CELL_SETTINGS.uiSimulationTimeFactor > UINT#100) THEN
	GVL_CELL_SETTINGS.uiSimulationTimeFactor := UINT#100;
END_IF;

// FB_AXIS являются единственными владельцами MC_Power. Группа получает только
// подтверждение готовности физических осей и управляет состоянием GroupStandby.
xDrivesPowered := GVL_AXIS.arrAxis[1].Status.xPowered
	AND GVL_AXIS.arrAxis[2].Status.xPowered
	AND GVL_AXIS.arrAxis[3].Status.xPowered;
lrGroupVelocityOverride := REAL_TO_LREAL(GVL_HMI.rRobotManualSpeedPercent) / 100.0;
IF xPointCheckActive THEN
	// Скорость проверки уже применяется FB_MOTION_MANAGER как VelFactor.
	// Глобальный override оставляем 100 %, иначе процент умножится сам на себя.
	lrGroupVelocityOverride := 1.0;
END_IF;
GVL_AXIS_GROUP.AxisGroup.MotionParam.HaltDeceleration := GVL_CELL_SETTINGS.lrRobotHaltDeceleration;
GVL_AXIS_GROUP.AxisGroup.MotionParam.HaltJerk := GVL_CELL_SETTINGS.lrRobotHaltJerk;
GROUP_XYZ(
	FaultRequest := stAxisGroupFaultRequest,
	xResetPermit := xRobotHmiPermit,
	xAxesPowered := xDrivesPowered,
	lrVelocityOverride := lrGroupVelocityOverride,
	AxisGroup := AXIS_GROUP_XYZ,
	GroupData := GVL_AXIS_GROUP.AxisGroup
);

// Повторная выборка после вызова FB публикует фактическое состояние текущего цикла.
xDrivesPowered := GVL_AXIS.arrAxis[1].Status.xPowered
	AND GVL_AXIS.arrAxis[2].Status.xPowered
	AND GVL_AXIS.arrAxis[3].Status.xPowered;
xAnyDrivePowered := GVL_AXIS.arrAxis[1].Status.xPowerStageOn
	OR GVL_AXIS.arrAxis[1].Status.xDriveStartOn
	OR GVL_AXIS.arrAxis[2].Status.xPowerStageOn
	OR GVL_AXIS.arrAxis[2].Status.xDriveStartOn
	OR GVL_AXIS.arrAxis[3].Status.xPowerStageOn
	OR GVL_AXIS.arrAxis[3].Status.xDriveStartOn;
xDrivesOff := NOT xAnyDrivePowered
	AND (GVL_AXIS_GROUP.AxisGroup.Diag.iStep = E_AXIS_GROUP_STATE.DISABLED);
xPowerTransitionActive :=
	(GVL_AXIS.arrAxis[1].Diag.iStep = E_AXIS_STATE.POWERING)
	OR (GVL_AXIS.arrAxis[1].Diag.iStep = E_AXIS_STATE.POWERING_DOWN)
	OR (GVL_AXIS.arrAxis[2].Diag.iStep = E_AXIS_STATE.POWERING)
	OR (GVL_AXIS.arrAxis[2].Diag.iStep = E_AXIS_STATE.POWERING_DOWN)
	OR (GVL_AXIS.arrAxis[3].Diag.iStep = E_AXIS_STATE.POWERING)
	OR (GVL_AXIS.arrAxis[3].Diag.iStep = E_AXIS_STATE.POWERING_DOWN)
	OR (GVL_AXIS_GROUP.AxisGroup.Diag.iStep = E_AXIS_GROUP_STATE.ENABLING_POWER)
	OR (GVL_AXIS_GROUP.AxisGroup.Diag.iStep = E_AXIS_GROUP_STATE.ENABLING_GROUP)
	OR (GVL_AXIS_GROUP.AxisGroup.Diag.iStep = E_AXIS_GROUP_STATE.DISABLING_GROUP)
	OR (GVL_AXIS_GROUP.AxisGroup.Diag.iStep = E_AXIS_GROUP_STATE.DISABLING_POWER);
xDrivesReady := GVL_AXIS.arrAxis[1].Status.xPowered
	AND GVL_AXIS.arrAxis[1].Status.xCanStartMotion
	AND NOT GVL_AXIS.arrAxis[1].Status.xError
	AND GVL_AXIS.arrAxis[2].Status.xPowered
	AND GVL_AXIS.arrAxis[2].Status.xCanStartMotion
	AND NOT GVL_AXIS.arrAxis[2].Status.xError
	AND GVL_AXIS.arrAxis[3].Status.xPowered
	AND GVL_AXIS.arrAxis[3].Status.xCanStartMotion
	AND NOT GVL_AXIS.arrAxis[3].Status.xError
	AND (GVL_AXIS_GROUP.AxisGroup.Diag.iStep = E_AXIS_GROUP_STATE.READY)
	AND NOT GVL_AXIS_GROUP.AxisGroup.Status.xLocalError
	AND NOT GVL_AXIS_GROUP.AxisGroup.Status.xLogicalError
	AND NOT GVL_AXIS_GROUP.AxisGroup.Status.xGroupError
	AND NOT SIMULATION_DYNAMICS.xBusy
	AND NOT SIMULATION_DYNAMICS.xError;
xAxisDriveError := GVL_AXIS.arrAxis[1].Status.xAxisError
	OR GVL_AXIS.arrAxis[1].Status.xLogicalError
	OR GVL_AXIS.arrAxis[2].Status.xAxisError
	OR GVL_AXIS.arrAxis[2].Status.xLogicalError
	OR GVL_AXIS.arrAxis[3].Status.xAxisError
	OR GVL_AXIS.arrAxis[3].Status.xLogicalError;
xGroupError := GVL_AXIS_GROUP.AxisGroup.Status.xLocalError
	OR GVL_AXIS_GROUP.AxisGroup.Status.xLogicalError
	OR GVL_AXIS_GROUP.AxisGroup.Status.xGroupError;
xDriveError := xAxisDriveError OR xGroupError;
xGroupMotionBusy := GVL_AXIS_GROUP.AxisGroup.Command.xMoveDirect
	OR GVL_AXIS_GROUP.AxisGroup.Command.xMoveLinear
	OR (GVL_AXIS_GROUP.AxisGroup.Diag.iStep = E_AXIS_GROUP_STATE.MOVING_DIRECT)
	OR (GVL_AXIS_GROUP.AxisGroup.Diag.iStep = E_AXIS_GROUP_STATE.MOVING_LINEAR)
	OR (GVL_AXIS_GROUP.AxisGroup.Diag.iStep = E_AXIS_GROUP_STATE.EMG_STOP)
	OR (GVL_AXIS_GROUP.AxisGroup.Diag.iStep = E_AXIS_GROUP_STATE.HALT_STOP)
	OR (GVL_AXIS_GROUP.AxisGroup.Diag.iStep = E_AXIS_GROUP_STATE.WAIT_STOP);
xMotionBusy := GVL_AXIS.arrAxis[1].Status.xMotionBusy
	OR GVL_AXIS.arrAxis[2].Status.xMotionBusy
	OR GVL_AXIS.arrAxis[3].Status.xMotionBusy
	OR xGroupMotionBusy;

// Повторно определяем владельца после вызова FB: на этом этапе уже виден
// переход READY -> HOMING/MOVE/JOG, даже если Motion FB станет Busy позже.
uiManualAxisOwner := UINT#0;
FOR uiMachine := 1 TO 3 DO
	IF (uiManualAxisOwner = UINT#0)
	AND (GVL_AXIS.arrAxis[uiMachine].Status.xMotionBusy
		OR (GVL_AXIS.arrAxis[uiMachine].Diag.iStep = E_AXIS_STATE.JOGGING)
		OR (GVL_AXIS.arrAxis[uiMachine].Diag.iStep = E_AXIS_STATE.JOG_DECELERATING)
		OR (GVL_AXIS.arrAxis[uiMachine].Diag.iStep = E_AXIS_STATE.HOMING)
		OR (GVL_AXIS.arrAxis[uiMachine].Diag.iStep = E_AXIS_STATE.MOVE_ABSOLUTE)
		OR (GVL_AXIS.arrAxis[uiMachine].Diag.iStep = E_AXIS_STATE.MOVE_RELATIVE)
		OR (GVL_AXIS.arrAxis[uiMachine].Diag.iStep = E_AXIS_STATE.STOPPING)
		OR (GVL_AXIS.arrAxis[uiMachine].Diag.iStep = E_AXIS_STATE.STOP_RELEASE)) THEN
		uiManualAxisOwner := uiMachine;
	END_IF;
END_FOR;
xMotionBusy := xMotionBusy OR (uiManualAxisOwner > UINT#0);

GVL_HMI.stRobotHmiStatus.xDrivesPowered := xDrivesPowered;
GVL_HMI.stRobotHmiStatus.xDrivesOff := xDrivesOff;
GVL_HMI.stRobotHmiStatus.xPowerTransitionActive := xPowerTransitionActive;
GVL_HMI.stRobotHmiStatus.xDrivesEnableAllowed := xRobotHmiPermit
	AND xHmiConnectionAlive
	AND NOT GVL_HMI.xModbusMode
	AND (NOT GVL_CELL_CONTROL.xGlobalError OR xManualRecoveryActive)
	AND xDrivesOff
	AND NOT xAxisDriveError
	AND NOT xRobotMotionCommandActive
	AND NOT xMotionBusy
	AND NOT xMotionResetBusy;
GVL_HMI.stRobotHmiStatus.xDrivesDisableAllowed := xRobotHmiPermit
	AND xHmiConnectionAlive
	AND NOT GVL_HMI.xModbusMode
	AND (xAnyDrivePowered
		OR (GVL_AXIS_GROUP.AxisGroup.Diag.iStep = E_AXIS_GROUP_STATE.READY))
	AND NOT xPowerTransitionActive
	AND NOT xRobotMotionCommandActive
	AND NOT xMotionBusy
	AND NOT xMotionResetBusy;
GVL_HMI.stRobotHmiStatus.xResetAllowed := xRobotHmiPermit
	AND xHmiConnectionAlive
	AND NOT GVL_HMI.xModbusMode
	AND (NOT GVL_CELL_CONTROL.xGlobalError OR xManualRecoveryActive)
	AND NOT xMotionBusy
	AND NOT xMotionResetBusy;
GVL_HMI.stRobotHmiStatus.xStopAllowed := xRobotHmiPermit
	AND xHmiConnectionAlive
	AND NOT GVL_HMI.xModbusMode
	AND (xMotionBusy OR xRobotMotionCommandActive);

// Финальная публикация разрешений выполняется после всех Motion FB. HMI получает
// актуальные статусы текущего цикла и не дублирует технологические условия.
FOR uiMachine := 1 TO 3 DO
	GVL_HMI.astAxisHmiStatus[uiMachine].lrActualPosition := GVL_AXIS.arrAxis[uiMachine].Status.lrActualPosition;
	GVL_HMI.astAxisHmiStatus[uiMachine].lrTargetPosition := GVL_HMI.astAxisHmiCommand[uiMachine].lrTargetPosition;
	GVL_HMI.astAxisHmiStatus[uiMachine].lrDeviation :=
		GVL_HMI.astAxisHmiStatus[uiMachine].lrActualPosition
		- GVL_HMI.astAxisHmiStatus[uiMachine].lrTargetPosition;
	GVL_HMI.astAxisHmiStatus[uiMachine].xDriveReady := GVL_AXIS.arrAxis[uiMachine].Status.xPowered
		AND NOT GVL_AXIS.arrAxis[uiMachine].Status.xAxisError
		AND NOT GVL_AXIS.arrAxis[uiMachine].Status.xLogicalError;
	GVL_HMI.astAxisHmiStatus[uiMachine].xBusy := GVL_AXIS.arrAxis[uiMachine].Status.xMotionBusy
		OR (uiManualAxisOwner = uiMachine);
	GVL_HMI.astAxisHmiStatus[uiMachine].xError := GVL_AXIS.arrAxis[uiMachine].Status.xAxisError
		OR GVL_AXIS.arrAxis[uiMachine].Status.xLogicalError;
	GVL_HMI.astAxisHmiStatus[uiMachine].xHomed := GVL_AXIS.arrAxis[uiMachine].Status.xHomed;
	GVL_HMI.astAxisHmiStatus[uiMachine].lrCommandVelocity := alrRobotManualRatedVelocity[uiMachine]
		* REAL_TO_LREAL(rRobotManualEffectiveSpeedPercent) / 100.0;
	GVL_HMI.astAxisHmiStatus[uiMachine].lrMaxVelocity := alrRobotManualRatedVelocity[uiMachine];
	GVL_HMI.astAxisHmiStatus[uiMachine].eState := GVL_AXIS.arrAxis[uiMachine].Diag.iStep;

	axManualAxisBaseAllowed[uiMachine] := xRobotHmiPermit
		AND NOT GVL_TWO_PALLET.astStatus[1].xBusy AND NOT GVL_TWO_PALLET.astStatus[2].xBusy
		AND xHmiConnectionAlive
		AND NOT GVL_HMI.xModbusMode
		AND (NOT GVL_CELL_CONTROL.xGlobalError OR xManualRecoveryActive)
		AND NOT xDriveError
		AND NOT GVL_ROBOT.Status.xBusy
		AND (GVL_AXIS_GROUP.AxisGroup.Diag.iStep = E_AXIS_GROUP_STATE.READY)
		AND (NOT xMotionBusy OR (uiManualAxisOwner = uiMachine))
		AND GVL_AXIS.arrAxis[uiMachine].Status.xPowered
		AND NOT GVL_AXIS.arrAxis[uiMachine].Status.xAxisError
		AND NOT GVL_AXIS.arrAxis[uiMachine].Status.xLogicalError
		AND (
			((GVL_AXIS.arrAxis[uiMachine].Diag.iStep = E_AXIS_STATE.READY)
				AND GVL_AXIS.arrAxis[uiMachine].Status.xCanStartMotion)
			OR ((uiManualAxisOwner = uiMachine)
				AND ((GVL_AXIS.arrAxis[uiMachine].Diag.iStep = E_AXIS_STATE.JOGGING)
					OR (GVL_AXIS.arrAxis[uiMachine].Diag.iStep = E_AXIS_STATE.JOG_DECELERATING)))
		);

	GVL_HMI.astAxisHmiStatus[uiMachine].xJogPositiveAllowed := axManualAxisBaseAllowed[uiMachine]
		AND GVL_HMI.xRobotContinuousMode;
	GVL_HMI.astAxisHmiStatus[uiMachine].xJogNegativeAllowed := axManualAxisBaseAllowed[uiMachine]
		AND GVL_HMI.xRobotContinuousMode;
	GVL_HMI.astAxisHmiStatus[uiMachine].xHomeAllowed := axManualAxisBaseAllowed[uiMachine]
		AND NOT GVL_CELL_CONTROL.xGlobalError
		AND NOT xMotionBusy
		AND GVL_AXIS.arrAxis[uiMachine].Status.xCanStartMotion;
	GVL_HMI.astAxisHmiStatus[uiMachine].xMoveAbsoluteAllowed := axManualAxisBaseAllowed[uiMachine]
		AND NOT GVL_CELL_CONTROL.xGlobalError
		AND GVL_AXIS.arrAxis[uiMachine].Status.xHomed
		AND GVL_AXIS.arrAxis[uiMachine].Status.xCanStartMotion
		AND (GVL_HMI.astAxisHmiCommand[uiMachine].lrTargetPosition
			>= GVL_HMI.astAxisHmiStatus[uiMachine].lrMinPosition)
		AND (GVL_HMI.astAxisHmiCommand[uiMachine].lrTargetPosition
			<= GVL_HMI.astAxisHmiStatus[uiMachine].lrMaxPosition)
		AND (NOT axRobotSoftwareLimitsEnabled[uiMachine]
			OR (GVL_HMI.astAxisHmiCommand[uiMachine].lrTargetPosition
				>= alrRobotSoftwareMinPosition[uiMachine]))
		AND (NOT axRobotSoftwareLimitsEnabled[uiMachine]
			OR (GVL_HMI.astAxisHmiCommand[uiMachine].lrTargetPosition
				<= alrRobotSoftwareMaxPosition[uiMachine]));
	GVL_HMI.astAxisHmiStatus[uiMachine].xMoveRelativePositiveAllowed := axManualAxisBaseAllowed[uiMachine]
		AND NOT GVL_HMI.xRobotContinuousMode
		AND NOT GVL_CELL_CONTROL.xGlobalError
		AND GVL_AXIS.arrAxis[uiMachine].Status.xHomed
		AND GVL_AXIS.arrAxis[uiMachine].Status.xCanStartMotion
		AND (GVL_HMI.astAxisHmiStatus[uiMachine].lrActualPosition + GVL_HMI.lrRobotManualStep
			<= GVL_HMI.astAxisHmiStatus[uiMachine].lrMaxPosition)
		AND (NOT axRobotSoftwareLimitsEnabled[uiMachine]
			OR (GVL_HMI.astAxisHmiStatus[uiMachine].lrActualPosition + GVL_HMI.lrRobotManualStep
				<= alrRobotSoftwareMaxPosition[uiMachine]));
	GVL_HMI.astAxisHmiStatus[uiMachine].xMoveRelativeNegativeAllowed := axManualAxisBaseAllowed[uiMachine]
		AND NOT GVL_HMI.xRobotContinuousMode
		AND NOT GVL_CELL_CONTROL.xGlobalError
		AND GVL_AXIS.arrAxis[uiMachine].Status.xHomed
		AND GVL_AXIS.arrAxis[uiMachine].Status.xCanStartMotion
		AND (GVL_HMI.astAxisHmiStatus[uiMachine].lrActualPosition - GVL_HMI.lrRobotManualStep
			>= GVL_HMI.astAxisHmiStatus[uiMachine].lrMinPosition)
		AND (NOT axRobotSoftwareLimitsEnabled[uiMachine]
			OR (GVL_HMI.astAxisHmiStatus[uiMachine].lrActualPosition - GVL_HMI.lrRobotManualStep
				>= alrRobotSoftwareMinPosition[uiMachine]));

	IF NOT xHmiConnectionAlive THEN
		GVL_HMI.astAxisHmiStatus[uiMachine].eRejectReason := E_HMI_MANUAL_REJECT.HMI_OFFLINE;
	ELSIF NOT xRobotHmiPermit THEN
		GVL_HMI.astAxisHmiStatus[uiMachine].eRejectReason := E_HMI_MANUAL_REJECT.MANUAL_MODE_REQUIRED;
	ELSIF GVL_HMI.xModbusMode THEN
		GVL_HMI.astAxisHmiStatus[uiMachine].eRejectReason := E_HMI_MANUAL_REJECT.MODBUS_ACTIVE;
	ELSIF xDriveError THEN
		GVL_HMI.astAxisHmiStatus[uiMachine].eRejectReason := E_HMI_MANUAL_REJECT.DRIVE_ERROR;
	ELSIF NOT GVL_HMI.astAxisHmiStatus[uiMachine].xDriveReady THEN
		GVL_HMI.astAxisHmiStatus[uiMachine].eRejectReason := E_HMI_MANUAL_REJECT.DRIVES_DISABLED;
	ELSIF GVL_CELL_CONTROL.xGlobalError THEN
		GVL_HMI.astAxisHmiStatus[uiMachine].eRejectReason := E_HMI_MANUAL_REJECT.GLOBAL_ERROR_JOG_ONLY;
	ELSIF GVL_ROBOT.Status.xBusy THEN
		GVL_HMI.astAxisHmiStatus[uiMachine].eRejectReason := E_HMI_MANUAL_REJECT.ROBOT_BUSY;
	ELSIF xMotionBusy AND (uiManualAxisOwner <> uiMachine) THEN
		GVL_HMI.astAxisHmiStatus[uiMachine].eRejectReason := E_HMI_MANUAL_REJECT.AXIS_BUSY;
	ELSIF (GVL_AXIS_GROUP.AxisGroup.Diag.iStep <> E_AXIS_GROUP_STATE.READY) THEN
		GVL_HMI.astAxisHmiStatus[uiMachine].eRejectReason := E_HMI_MANUAL_REJECT.MOTION_NOT_READY;
	ELSIF NOT (
		((GVL_AXIS.arrAxis[uiMachine].Diag.iStep = E_AXIS_STATE.READY)
			AND GVL_AXIS.arrAxis[uiMachine].Status.xCanStartMotion)
		OR ((uiManualAxisOwner = uiMachine)
			AND ((GVL_AXIS.arrAxis[uiMachine].Diag.iStep = E_AXIS_STATE.JOGGING)
				OR (GVL_AXIS.arrAxis[uiMachine].Diag.iStep = E_AXIS_STATE.JOG_DECELERATING)))
	) THEN
		GVL_HMI.astAxisHmiStatus[uiMachine].eRejectReason := E_HMI_MANUAL_REJECT.MOTION_NOT_READY;
	ELSIF NOT GVL_HMI.xRobotContinuousMode
	AND NOT GVL_HMI.astAxisHmiStatus[uiMachine].xHomed THEN
		GVL_HMI.astAxisHmiStatus[uiMachine].eRejectReason := E_HMI_MANUAL_REJECT.AXIS_NOT_HOMED;
	ELSIF axManualAxisCommandRejected[uiMachine] THEN
		GVL_HMI.astAxisHmiStatus[uiMachine].eRejectReason := E_HMI_MANUAL_REJECT.COMMAND_CONFLICT;
	ELSE
		GVL_HMI.astAxisHmiStatus[uiMachine].eRejectReason := E_HMI_MANUAL_REJECT.NONE;
	END_IF;
END_FOR;

// PLC хранит владельца до фактического окончания торможения. Только после этого
// следующая мобильная аренда сможет получить новый фронт xMobileMotionActive.
IF xMobileMotionLeaseActive
AND NOT GVL_HMI.xMobileMotionActive
AND NOT xMotionBusy THEN
	xMobileMotionLeaseActive := FALSE;
	xMobileMotionStopRequest := FALSE;
	xMobileMotionConnectionAlive := FALSE;
	GVL_HMI.xMobileMotionLeaseAlive := FALSE;
END_IF;

IF NOT GVL_HMI.xModbusMode THEN
	GVL_HMI.lrActualX := GVL_AXIS_GROUP.AxisGroup.Status.ActualX;
	GVL_HMI.lrActualY := GVL_AXIS_GROUP.AxisGroup.Status.ActualY;
	GVL_HMI.lrActualZ := GVL_AXIS_GROUP.AxisGroup.Status.ActualZ;
	GVL_HMI.HMI.ActualX := GVL_HMI.lrActualX;
	GVL_HMI.HMI.ActualY := GVL_HMI.lrActualY;
	GVL_HMI.HMI.ActualZ := GVL_HMI.lrActualZ;
END_IF;
END_METHOD

METHOD PRIVATE RunGeometryControl
xGeometryEnvironmentChanged := NOT xGeometryInitialized
	OR (eGeometryPreviousEnvironment <> GVL_CELL_SETTINGS.eTestEnvironment);
GVL_GEOMETRY_CONTROL.uiEnvironment := TO_UINT(GVL_CELL_SETTINGS.eTestEnvironment);
GVL_GEOMETRY_CONTROL.xSupported := NOT GVL_HMI.xModbusMode
	AND (GVL_CELL_SETTINGS.eTestEnvironment <> E_CELL_TEST_ENVIRONMENT.SC500_BENCH);
IF xGeometryEnvironmentChanged THEN
	FOR uiGeometry := UINT#1 TO UINT#2 DO
		IF GVL_CELL_SETTINGS.eTestEnvironment = E_CELL_TEST_ENVIRONMENT.NORMAL THEN
			GVL_GEOMETRY_CONTROL.astActiveMemory[uiGeometry] := GVL_GEOMETRY_CONTROL.astMemory[uiGeometry];
		ELSE GVL_GEOMETRY_CONTROL.astActiveMemory[uiGeometry] := GVL_GEOMETRY_CONTROL.astSimulationMemory[uiGeometry]; END_IF;
		GVL_GEOMETRY_CONTROL.astSignals[uiGeometry].xReserve := FALSE;
		GVL_GEOMETRY_CONTROL.astSignals[uiGeometry].xDeposited := FALSE;
		GVL_GEOMETRY_CONTROL.astSignals[uiGeometry].xReleased := FALSE;
		GVL_GEOMETRY_CONTROL.astSignals[uiGeometry].xRobotInteraction := FALSE;
	END_FOR;
	FOR uiGeometryMachine := UINT#1 TO UINT#3 DO
		IF GVL_CELL_SETTINGS.eTestEnvironment = E_CELL_TEST_ENVIRONMENT.NORMAL THEN
			GVL_GEOMETRY_CONTROL.astCalls[uiGeometryMachine] := GVL_GEOMETRY_CONTROL.astRetainCalls[uiGeometryMachine];
			GVL_GEOMETRY_CONTROL.auiActiveCount[uiGeometryMachine] := GVL_GEOMETRY_CONTROL.auiCount[uiGeometryMachine];
		ELSE
			GVL_GEOMETRY_CONTROL.astCalls[uiGeometryMachine] := GVL_GEOMETRY_CONTROL.astSimulationCalls[uiGeometryMachine];
			GVL_GEOMETRY_CONTROL.auiActiveCount[uiGeometryMachine] := GVL_GEOMETRY_CONTROL.auiSimulationCount[uiGeometryMachine];
		END_IF;
		IF (GVL_GEOMETRY_CONTROL.astCalls[uiGeometryMachine].uiState = UINT#2)
		OR (GVL_GEOMETRY_CONTROL.astCalls[uiGeometryMachine].uiState = UINT#3) THEN
			GVL_GEOMETRY_CONTROL.astCalls[uiGeometryMachine].uiState := UINT#7;
			GVL_GEOMETRY_CONTROL.astCalls[uiGeometryMachine].uiReason := UINT#5;
			F_GEOMETRY_EVENT(Call := GVL_GEOMETRY_CONTROL.astCalls[uiGeometryMachine]);
		END_IF;
	END_FOR;
	xGeometryInitialized := TRUE;
	eGeometryPreviousEnvironment := GVL_CELL_SETTINGS.eTestEnvironment;
END_IF;
FOR uiGeometry := UINT#1 TO UINT#2 DO
	GVL_GEOMETRY_CONTROL.auiAction[uiGeometry] := UINT#0;
	IF GVL_CELL_SETTINGS.eTestEnvironment = E_CELL_TEST_ENVIRONMENT.NORMAL THEN
		GVL_GEOMETRY_CONTROL.astActiveConfig[uiGeometry] := GVL_GEOMETRY_CONTROL.astConfig[uiGeometry];
	ELSE GVL_GEOMETRY_CONTROL.astActiveConfig[uiGeometry] := GVL_GEOMETRY_CONTROL.astSimulationConfig[uiGeometry]; END_IF;
END_FOR;
GVL_GEOMETRY_CONTROL.xAutoChangeAllowed := GVL_GEOMETRY_CONTROL.xSupported
	AND xHmiConnectionAlive AND NOT GVL_HMI.xTestSessionActive AND NOT GVL_CELL_CONTROL.xGlobalError;
GVL_GEOMETRY_CONTROL.xSettingsAllowed := GVL_GEOMETRY_CONTROL.xSupported
	AND GVL_CELL_SETTINGS.xCellSettingsChangeAllowed AND xHmiConnectionAlive
	AND NOT GVL_GEOMETRY_CONTROL.astStatus[1].xDriveRunning AND NOT GVL_GEOMETRY_CONTROL.astStatus[2].xDriveRunning
	AND NOT GVL_GEOMETRY_CONTROL.astStatus[1].xResetBusy AND NOT GVL_GEOMETRY_CONTROL.astStatus[2].xResetBusy
	AND NOT GVL_GEOMETRY_CONTROL.astStatus[1].xReserved AND NOT GVL_GEOMETRY_CONTROL.astStatus[2].xReserved
	AND NOT GVL_GEOMETRY_CONTROL.astSignals[1].xRobotInteraction AND NOT GVL_GEOMETRY_CONTROL.astSignals[2].xRobotInteraction
	AND NOT GEOMETRY[1].xRunOutput AND NOT GEOMETRY[2].xRunOutput;
FOR uiGeometryMachine := UINT#1 TO UINT#3 DO
	GVL_GEOMETRY_CONTROL.axCallAllowed[uiGeometryMachine] := GVL_GEOMETRY_CONTROL.xAutoChangeAllowed
		AND GVL_MACHINE.Status[uiGeometryMachine].xEnabled
		AND ((GVL_GEOMETRY_CONTROL.astCalls[uiGeometryMachine].uiState <= UINT#1)
			OR (GVL_GEOMETRY_CONTROL.astCalls[uiGeometryMachine].uiState > UINT#3))
		AND (GVL_GEOMETRY_CONTROL.astStatus[1].xEnabled OR GVL_GEOMETRY_CONTROL.astStatus[2].xEnabled);
	GVL_GEOMETRY_CONTROL.axCancelAllowed[uiGeometryMachine] := GVL_GEOMETRY_CONTROL.xAutoChangeAllowed
		AND (GVL_GEOMETRY_CONTROL.astCalls[uiGeometryMachine].uiState = UINT#1);
END_FOR;

